    #Ok := "FRK_ConfigDecode"(Text := STRING_TO_WSTRING("FRK_PersistImages".D010.Rows[6].Record.ValueText), Storage := 3, Minimum := 0.0, Maximum := 1000.0, MaxLength := 0, Value := "FRK_ConfigScratch".Value);
    IF NOT #Ok THEN RETURN; END_IF;
    IF NOT "FRK_PersistImages".D010.Rows[7].Used OR "FRK_PersistImages".D010.Rows[7].SchemaVersion <> 4 OR "FRK_PersistImages".D010.Rows[7].ModelCode <> 'MODEL_A' OR "FRK_PersistImages".D010.Rows[7].Record.Scope <> 'StationB.Cell.Gate' OR "FRK_PersistImages".D010.Rows[7].Record.WriteKey <> 'timeout' OR "FRK_PersistImages".D010.Rows[7].Record.Revision <> 1 OR "FRK_PersistImages".D010.Rows[7].Record.Kind <> 0 OR "FRK_PersistImages".D010.Rows[7].Record.ValueType <> 3 THEN RETURN; END_IF;
    #Ok := "FRK_ConfigDecode"(Text := STRING_TO_WSTRING("FRK_PersistImages".D010.Rows[7].Record.ValueText), Storage := 7, Minimum := 1.0, Maximum := 60000.0, MaxLength := 0, Value := "FRK_ConfigScratch".Value);
    IF NOT #Ok THEN RETURN; END_IF;
    IF NOT "FRK_PersistImages".D010.Rows[8].Used OR "FRK_PersistImages".D010.Rows[8].SchemaVersion <> 4 OR "FRK_PersistImages".D010.Rows[8].ModelCode <> 'MODEL_A' OR "FRK_PersistImages".D010.Rows[8].Record.Scope <> 'StationB.Cell.Gate' OR "FRK_PersistImages".D010.Rows[8].Record.WriteKey <> 'preset' OR "FRK_PersistImages".D010.Rows[8].Record.Revision <> 2 OR "FRK_PersistImages".D010.Rows[8].Record.Kind <> 0 OR "FRK_PersistImages".D010.Rows[8].Record.ValueType <> 0 THEN RETURN; END_IF;
    #Ok := "FRK_ConfigDecode"(Text := STRING_TO_WSTRING("FRK_PersistImages".D010.Rows[8].Record.ValueText), Storage := 3, Minimum := 0.0, Maximum := 1000.0, MaxLength := 0, Value := "FRK_ConfigScratch".Value);
    IF NOT #Ok THEN RETURN; END_IF;
    IF NOT "FRK_PersistImages".D010.Rows[9].Used OR "FRK_PersistImages".D010.Rows[9].SchemaVersion <> 4 OR "FRK_PersistImages".D010.Rows[9].ModelCode <> 'MODEL_A' OR "FRK_PersistImages".D010.Rows[9].Record.Scope <> 'StationB.Satellite' OR "FRK_PersistImages".D010.Rows[9].Record.WriteKey <> 'timeout' OR "FRK_PersistImages".D010.Rows[9].Record.Revision <> 1 OR "FRK_PersistImages".D010.Rows[9].Record.Kind <> 0 OR "FRK_PersistImages".D010.Rows[9].Record.ValueType <> 3 THEN RETURN; END_IF;
    #Ok := "FRK_ConfigDecode"(Text := STRING_TO_WSTRING("FRK_PersistImages".D010.Rows[9].Record.ValueText), Storage := 7, Minimum := 1.0, Maximum := 60000.0, MaxLength := 0, Value := "FRK_ConfigScratch".Value);
    IF NOT #Ok THEN RETURN; END_IF;
    IF NOT "FRK_PersistImages".D010.Rows[10].Used OR "FRK_PersistImages".D010.Rows[10].SchemaVersion <> 4 OR "FRK_PersistImages".D010.Rows[10].ModelCode <> 'MODEL_A' OR "FRK_PersistImages".D010.Rows[10].Record.Scope <> 'StationB.Satellite' OR "FRK_PersistImages".D010.Rows[10].Record.WriteKey <> 'preset' OR "FRK_PersistImages".D010.Rows[10].Record.Revision <> 2 OR "FRK_PersistImages".D010.Rows[10].Record.Kind <> 0 OR "FRK_PersistImages".D010.Rows[10].Record.ValueType <> 0 THEN RETURN; END_IF;
    #Ok := "FRK_ConfigDecode"(Text := STRING_TO_WSTRING("FRK_PersistImages".D010.Rows[10].Record.ValueText), Storage := 3, Minimum := 0.0, Maximum := 1000.0, MaxLength := 0, Value := "FRK_ConfigScratch".Value);
    IF NOT #Ok THEN RETURN; END_IF;
    IF NOT "FRK_PersistImages".D010.Rows[11].Used OR "FRK_PersistImages".D010.Rows[11].SchemaVersion <> 4 OR "FRK_PersistImages".D010.Rows[11].ModelCode <> 'MODEL_A' OR "FRK_PersistImages".D010.Rows[11].Record.Scope <> 'StationB.Satellite.Cell' OR "FRK_PersistImages".D010.Rows[11].Record.WriteKey <> 'timeout' OR "FRK_PersistImages".D010.Rows[11].Record.Revision <> 1 OR "FRK_PersistImages".D010.Rows[11].Record.Kind <> 0 OR "FRK_PersistImages".D010.Rows[11].Record.ValueType <> 3 THEN RETURN; END_IF;
    #Ok := "FRK_ConfigDecode"(Text := STRING_TO_WSTRING("FRK_PersistImages".D010.Rows[11].Record.ValueText), Storage := 7, Minimum := 1.0, Maximum := 60000.0, MaxLength := 0, Value := "FRK_ConfigScratch".Value);
    IF NOT #Ok THEN RETURN; END_IF;
    IF NOT "FRK_PersistImages".D010.Rows[12].Used OR "FRK_PersistImages".D010.Rows[12].SchemaVersion <> 4 OR "FRK_PersistImages".D010.Rows[12].ModelCode <> 'MODEL_A' OR "FRK_PersistImages".D010.Rows[12].Record.Scope <> 'StationB.Satellite.Cell' OR "FRK_PersistImages".D010.Rows[12].Record.WriteKey <> 'preset' OR "FRK_PersistImages".D010.Rows[12].Record.Revision <> 2 OR "FRK_PersistImages".D010.Rows[12].Record.Kind <> 0 OR "FRK_PersistImages".D010.Rows[12].Record.ValueType <> 0 THEN RETURN; END_IF;
    #Ok := "FRK_ConfigDecode"(Text := STRING_TO_WSTRING("FRK_PersistImages".D010.Rows[12].Record.ValueText), Storage := 3, Minimum := 0.0, Maximum := 1000.0, MaxLength := 0, Value := "FRK_ConfigScratch".Value);
    IF NOT #Ok THEN RETURN; END_IF;
    IF NOT "FRK_PersistImages".D010.Rows[13].Used OR "FRK_PersistImages".D010.Rows[13].SchemaVersion <> 4 OR "FRK_PersistImages".D010.Rows[13].ModelCode <> 'MODEL_A' OR "FRK_PersistImages".D010.Rows[13].Record.Scope <> 'StationB.Satellite.Cell.Clamp' OR "FRK_PersistImages".D010.Rows[13].Record.WriteKey <> 'timeout' OR "FRK_PersistImages".D010.Rows[13].Record.Revision <> 1 OR "FRK_PersistImages".D010.Rows[13].Record.Kind <> 0 OR "FRK_PersistImages".D010.Rows[13].Record.ValueType <> 3 THEN RETURN; END_IF;
    #Ok := "FRK_ConfigDecode"(Text := STRING_TO_WSTRING("FRK_PersistImages".D010.Rows[13].Record.ValueText), Storage := 7, Minimum := 1.0, Maximum := 60000.0, MaxLength := 0, Value := "FRK_ConfigScratch".Value);
    IF NOT #Ok THEN RETURN; END_IF;
    IF NOT "FRK_PersistImages".D010.Rows[14].Used OR "FRK_PersistImages".D010.Rows[14].SchemaVersion <> 4 OR "FRK_PersistImages".D010.Rows[14].ModelCode <> 'MODEL_A' OR "FRK_PersistImages".D010.Rows[14].Record.Scope <> 'StationB.Satellite.Cell.Clamp' OR "FRK_PersistImages".D010.Rows[14].Record.WriteKey <> 'preset' OR "FRK_PersistImages".D010.Rows[14].Record.Revision <> 2 OR "FRK_PersistImages".D010.Rows[14].Record.Kind <> 0 OR "FRK_PersistImages".D010.Rows[14].Record.ValueType <> 0 THEN RETURN; END_IF;
    #Ok := "FRK_ConfigDecode"(Text := STRING_TO_WSTRING("FRK_PersistImages".D010.Rows[14].Record.ValueText), Storage := 3, Minimum := 0.0, Maximum := 1000.0, MaxLength := 0, Value := "FRK_ConfigScratch".Value);
    IF NOT #Ok THEN RETURN; END_IF;
    IF NOT "FRK_PersistImages".D010.Rows[15].Used OR "FRK_PersistImages".D010.Rows[15].SchemaVersion <> 4 OR "FRK_PersistImages".D010.Rows[15].ModelCode <> 'MODEL_A' OR "FRK_PersistImages".D010.Rows[15].Record.Scope <> 'StationB.Satellite.Cell.Gate' OR "FRK_PersistImages".D010.Rows[15].Record.WriteKey <> 'timeout' OR "FRK_PersistImages".D010.Rows[15].Record.Revision <> 1 OR "FRK_PersistImages".D010.Rows[15].Record.Kind <> 0 OR "FRK_PersistImages".D010.Rows[15].Record.ValueType <> 3 THEN RETURN; END_IF;
    #Ok := "FRK_ConfigDecode"(Text := STRING_TO_WSTRING("FRK_PersistImages".D010.Rows[15].Record.ValueText), Storage := 7, Minimum := 1.0, Maximum := 60000.0, MaxLength := 0, Value := "FRK_ConfigScratch".Value);
    IF NOT #Ok THEN RETURN; END_IF;
    IF NOT "FRK_PersistImages".D010.Rows[16].Used OR "FRK_PersistImages".D010.Rows[16].SchemaVersion <> 4 OR "FRK_PersistImages".D010.Rows[16].ModelCode <> 'MODEL_A' OR "FRK_PersistImages".D010.Rows[16].Record.Scope <> 'StationB.Satellite.Cell.Gate' OR "FRK_PersistImages".D010.Rows[16].Record.WriteKey <> 'preset' OR "FRK_PersistImages".D010.Rows[16].Record.Revision <> 2 OR "FRK_PersistImages".D010.Rows[16].Record.Kind <> 0 OR "FRK_PersistImages".D010.Rows[16].Record.ValueType <> 0 THEN RETURN; END_IF;
    #Ok := "FRK_ConfigDecode"(Text := STRING_TO_WSTRING("FRK_PersistImages".D010.Rows[16].Record.ValueText), Storage := 3, Minimum := 0.0, Maximum := 1000.0, MaxLength := 0, Value := "FRK_ConfigScratch".Value);
    IF NOT #Ok THEN RETURN; END_IF;
    IF NOT "FRK_PersistImages".D010.Rows[17].Used OR "FRK_PersistImages".D010.Rows[17].SchemaVersion <> 4 OR "FRK_PersistImages".D010.Rows[17].ModelCode <> 'MODEL_A' OR "FRK_PersistImages".D010.Rows[17].Record.Scope <> 'StationB.Satellite.Inner' OR "FRK_PersistImages".D010.Rows[17].Record.WriteKey <> 'timeout' OR "FRK_PersistImages".D010.Rows[17].Record.Revision <> 1 OR "FRK_PersistImages".D010.Rows[17].Record.Kind <> 0 OR "FRK_PersistImages".D010.Rows[17].Record.ValueType <> 3 THEN RETURN; END_IF;
    #Ok := "FRK_ConfigDecode"(Text := STRING_TO_WSTRING("FRK_PersistImages".D010.Rows[17].Record.ValueText), Storage := 7, Minimum := 1.0, Maximum := 60000.0, MaxLength := 0, Value := "FRK_ConfigScratch".Value);
    IF NOT #Ok THEN RETURN; END_IF;
    IF NOT "FRK_PersistImages".D010.Rows[18].Used OR "FRK_PersistImages".D010.Rows[18].SchemaVersion <> 4 OR "FRK_PersistImages".D010.Rows[18].ModelCode <> 'MODEL_A' OR "FRK_PersistImages".D010.Rows[18].Record.Scope <> 'StationB.Satellite.Inner' OR "FRK_PersistImages".D010.Rows[18].Record.WriteKey <> 'preset' OR "FRK_PersistImages".D010.Rows[18].Record.Revision <> 2 OR "FRK_PersistImages".D010.Rows[18].Record.Kind <> 0 OR "FRK_PersistImages".D010.Rows[18].Record.ValueType <> 0 THEN RETURN; END_IF;
    #Ok := "FRK_ConfigDecode"(Text := STRING_TO_WSTRING("FRK_PersistImages".D010.Rows[18].Record.ValueText), Storage := 3, Minimum := 0.0, Maximum := 1000.0, MaxLength := 0, Value := "FRK_ConfigScratch".Value);
    IF NOT #Ok THEN RETURN; END_IF;
    IF NOT "FRK_PersistImages".D010.Rows[19].Used OR "FRK_PersistImages".D010.Rows[19].SchemaVersion <> 4 OR "FRK_PersistImages".D010.Rows[19].ModelCode <> 'MODEL_A' OR "FRK_PersistImages".D010.Rows[19].Record.Scope <> 'StationB.Satellite.Inner.Cell' OR "FRK_PersistImages".D010.Rows[19].Record.WriteKey <> 'timeout' OR "FRK_PersistImages".D010.Rows[19].Record.Revision <> 1 OR "FRK_PersistImages".D010.Rows[19].Record.Kind <> 0 OR "FRK_PersistImages".D010.Rows[19].Record.ValueType <> 3 THEN RETURN; END_IF;
    #Ok := "FRK_ConfigDecode"(Text := STRING_TO_WSTRING("FRK_PersistImages".D010.Rows[19].Record.ValueText), Storage := 7, Minimum := 1.0, Maximum := 60000.0, MaxLength := 0, Value := "FRK_ConfigScratch".Value);
    IF NOT #Ok THEN RETURN; END_IF;
    IF NOT "FRK_PersistImages".D010.Rows[20].Used OR "FRK_PersistImages".D010.Rows[20].SchemaVersion <> 4 OR "FRK_PersistImages".D010.Rows[20].ModelCode <> 'MODEL_A' OR "FRK_PersistImages".D010.Rows[20].Record.Scope <> 'StationB.Satellite.Inner.Cell' OR "FRK_PersistImages".D010.Rows[20].Record.WriteKey <> 'preset' OR "FRK_PersistImages".D010.Rows[20].Record.Revision <> 2 OR "FRK_PersistImages".D010.Rows[20].Record.Kind <> 0 OR "FRK_PersistImages".D010.Rows[20].Record.ValueType <> 0 THEN RETURN; END_IF;
    #Ok := "FRK_ConfigDecode"(Text := STRING_TO_WSTRING("FRK_PersistImages".D010.Rows[20].Record.ValueText), Storage := 3, Minimum := 0.0, Maximum := 1000.0, MaxLength := 0, Value := "FRK_ConfigScratch".Value);
    IF NOT #Ok THEN RETURN; END_IF;
    IF NOT "FRK_PersistImages".D010.Rows[21].Used OR "FRK_PersistImages".D010.Rows[21].SchemaVersion <> 4 OR "FRK_PersistImages".D010.Rows[21].ModelCode <> 'MODEL_A' OR "FRK_PersistImages".D010.Rows[21].Record.Scope <> 'StationB.Satellite.Inner.Cell.Clamp' OR "FRK_PersistImages".D010.Rows[21].Record.WriteKey <> 'timeout' OR "FRK_PersistImages".D010.Rows[21].Record.Revision <> 1 OR "FRK_PersistImages".D010.Rows[21].Record.Kind <> 0 OR "FRK_PersistImages".D010.Rows[21].Record.ValueType <> 3 THEN RETURN; END_IF;
    #Ok := "FRK_ConfigDecode"(Text := STRING_TO_WSTRING("FRK_PersistImages".D010.Rows[21].Record.ValueText), Storage := 7, Minimum := 1.0, Maximum := 60000.0, MaxLength := 0, Value := "FRK_ConfigScratch".Value);
    IF NOT #Ok THEN RETURN; END_IF;
    IF NOT "FRK_PersistImages".D010.Rows[22].Used OR "FRK_PersistImages".D010.Rows[22].SchemaVersion <> 4 OR "FRK_PersistImages".D010.Rows[22].ModelCode <> 'MODEL_A' OR "FRK_PersistImages".D010.Rows[22].Record.Scope <> 'StationB.Satellite.Inner.Cell.Clamp' OR "FRK_PersistImages".D010.Rows[22].Record.WriteKey <> 'preset' OR "FRK_PersistImages".D010.Rows[22].Record.Revision <> 2 OR "FRK_PersistImages".D010.Rows[22].Record.Kind <> 0 OR "FRK_PersistImages".D010.Rows[22].Record.ValueType <> 0 THEN RETURN; END_IF;
    #Ok := "FRK_ConfigDecode"(Text := STRING_TO_WSTRING("FRK_PersistImages".D010.Rows[22].Record.ValueText), Storage := 3, Minimum := 0.0, Maximum := 1000.0, MaxLength := 0, Value := "FRK_ConfigScratch".Value);
    IF NOT #Ok THEN RETURN; END_IF;
    IF NOT "FRK_PersistImages".D010.Rows[23].Used OR "FRK_PersistImages".D010.Rows[23].SchemaVersion <> 4 OR "FRK_PersistImages".D010.Rows[23].ModelCode <> 'MODEL_A' OR "FRK_PersistImages".D010.Rows[23].Record.Scope <> 'StationB.Satellite.Inner.Cell.Gate' OR "FRK_PersistImages".D010.Rows[23].Record.WriteKey <> 'timeout' OR "FRK_PersistImages".D010.Rows[23].Record.Revision <> 1 OR "FRK_PersistImages".D010.Rows[23].Record.Kind <> 0 OR "FRK_PersistImages".D010.Rows[23].Record.ValueType <> 3 THEN RETURN; END_IF;
    #Ok := "FRK_ConfigDecode"(Text := STRING_TO_WSTRING("FRK_PersistImages".D010.Rows[23].Record.ValueText), Storage := 7, Minimum := 1.0, Maximum := 60000.0, MaxLength := 0, Value := "FRK_ConfigScratch".Value);
    IF NOT #Ok THEN RETURN; END_IF;
    IF NOT "FRK_PersistImages".D010.Rows[24].Used OR "FRK_PersistImages".D010.Rows[24].SchemaVersion <> 4 OR "FRK_PersistImages".D010.Rows[24].ModelCode <> 'MODEL_A' OR "FRK_PersistImages".D010.Rows[24].Record.Scope <> 'StationB.Satellite.Inner.Cell.Gate' OR "FRK_PersistImages".D010.Rows[24].Record.WriteKey <> 'preset' OR "FRK_PersistImages".D010.Rows[24].Record.Revision <> 2 OR "FRK_PersistImages".D010.Rows[24].Record.Kind <> 0 OR "FRK_PersistImages".D010.Rows[24].Record.ValueType <> 0 THEN RETURN; END_IF;
    #Ok := "FRK_ConfigDecode"(Text := STRING_TO_WSTRING("FRK_PersistImages".D010.Rows[24].Record.ValueText), Storage := 3, Minimum := 0.0, Maximum := 1000.0, MaxLength := 0, Value := "FRK_ConfigScratch".Value);
    IF NOT #Ok THEN RETURN; END_IF;
    #Stored := "FRK_ConfigFind"(Scope := 'StationB', Key := 'timeout', ModelCode := 'MODEL_A');
    IF #Stored = 0 THEN
        FOR #Index := 1 TO 114 DO
            #Reserved := NOT "FRK_ConfigStore".Rows[#Index].Used;
            FOR #Prior := 1 TO 0 DO IF #Targets[#Prior] = #Index THEN #Reserved := FALSE; END_IF; END_FOR;
            IF #Reserved THEN #Stored := #Index; EXIT; END_IF;
        END_FOR;
    END_IF;
    IF #Stored < 1 OR #Stored > 114 THEN RETURN; END_IF;
    #Targets[1] := #Stored;
    #Stored := "FRK_ConfigFind"(Scope := 'StationB', Key := 'preset', ModelCode := 'MODEL_A');
    IF #Stored = 0 THEN
        FOR #Index := 1 TO 114 DO
            #Reserved := NOT "FRK_ConfigStore".Rows[#Index].Used;
            FOR #Prior := 1 TO 1 DO IF #Targets[#Prior] = #Index THEN #Reserved := FALSE; END_IF; END_FOR;
            IF #Reserved THEN #Stored := #Index; EXIT; END_IF;
        END_FOR;
    END_IF;
    IF #Stored < 1 OR #Stored > 114 THEN RETURN; END_IF;
    #Targets[2] := #Stored;
    #Stored := "FRK_ConfigFind"(Scope := 'StationB.Cell', Key := 'timeout', ModelCode := 'MODEL_A');
    IF #Stored = 0 THEN
        FOR #Index := 1 TO 114 DO
            #Reserved := NOT "FRK_ConfigStore".Rows[#Index].Used;
            FOR #Prior := 1 TO 2 DO IF #Targets[#Prior] = #Index THEN #Reserved := FALSE; END_IF; END_FOR;
            IF #Reserved THEN #Stored := #Index; EXIT; END_IF;
        END_FOR;
    END_IF;
    IF #Stored < 1 OR #Stored > 114 THEN RETURN; END_IF;
    #Targets[3] := #Stored;
    #Stored := "FRK_ConfigFind"(Scope := 'StationB.Cell', Key := 'preset', ModelCode := 'MODEL_A');
    IF #Stored = 0 THEN
        FOR #Index := 1 TO 114 DO
            #Reserved := NOT "FRK_ConfigStore".Rows[#Index].Used;
            FOR #Prior := 1 TO 3 DO IF #Targets[#Prior] = #Index THEN #Reserved := FALSE; END_IF; END_FOR;
            IF #Reserved THEN #Stored := #Index; EXIT; END_IF;
        END_FOR;
    END_IF;
    IF #Stored < 1 OR #Stored > 114 THEN RETURN; END_IF;
    #Targets[4] := #Stored;
    #Stored := "FRK_ConfigFind"(Scope := 'StationB.Cell.Clamp', Key := 'timeout', ModelCode := 'MODEL_A');
    IF #Stored = 0 THEN
        FOR #Index := 1 TO 114 DO
            #Reserved := NOT "FRK_ConfigStore".Rows[#Index].Used;
            FOR #Prior := 1 TO 4 DO IF #Targets[#Prior] = #Index THEN #Reserved := FALSE; END_IF; END_FOR;
            IF #Reserved THEN #Stored := #Index; EXIT; END_IF;
        END_FOR;
    END_IF;
    IF #Stored < 1 OR #Stored > 114 THEN RETURN; END_IF;
    #Targets[5] := #Stored;
    #Stored := "FRK_ConfigFind"(Scope := 'StationB.Cell.Clamp', Key := 'preset', ModelCode := 'MODEL_A');
    IF #Stored = 0 THEN
        FOR #Index := 1 TO 114 DO
            #Reserved := NOT "FRK_ConfigStore".Rows[#Index].Used;
            FOR #Prior := 1 TO 5 DO IF #Targets[#Prior] = #Index THEN #Reserved := FALSE; END_IF; END_FOR;
            IF #Reserved THEN #Stored := #Index; EXIT; END_IF;
        END_FOR;
    END_IF;
    IF #Stored < 1 OR #Stored > 114 THEN RETURN; END_IF;
    #Targets[6] := #Stored;
    #Stored := "FRK_ConfigFind"(Scope := 'StationB.Cell.Gate', Key := 'timeout', ModelCode := 'MODEL_A');
    IF #Stored = 0 THEN
        FOR #Index := 1 TO 114 DO
            #Reserved := NOT "FRK_ConfigStore".Rows[#Index].Used;
            FOR #Prior := 1 TO 6 DO IF #Targets[#Prior] = #Index THEN #Reserved := FALSE; END_IF; END_FOR;
            IF #Reserved THEN #Stored := #Index; EXIT; END_IF;
        END_FOR;
    END_IF;
    IF #Stored < 1 OR #Stored > 114 THEN RETURN; END_IF;
    #Targets[7] := #Stored;
    #Stored := "FRK_ConfigFind"(Scope := 'StationB.Cell.Gate', Key := 'preset', ModelCode := 'MODEL_A');
    IF #Stored = 0 THEN
        FOR #Index := 1 TO 114 DO
            #Reserved := NOT "FRK_ConfigStore".Rows[#Index].Used;
            FOR #Prior := 1 TO 7 DO IF #Targets[#Prior] = #Index THEN #Reserved := FALSE; END_IF; END_FOR;
            IF #Reserved THEN #Stored := #Index; EXIT; END_IF;
        END_FOR;
    END_IF;
    IF #Stored < 1 OR #Stored > 114 THEN RETURN; END_IF;
    #Targets[8] := #Stored;
    #Stored := "FRK_ConfigFind"(Scope := 'StationB.Satellite', Key := 'timeout', ModelCode := 'MODEL_A');
    IF #Stored = 0 THEN
        FOR #Index := 1 TO 114 DO
            #Reserved := NOT "FRK_ConfigStore".Rows[#Index].Used;
            FOR #Prior := 1 TO 8 DO IF #Targets[#Prior] = #Index THEN #Reserved := FALSE; END_IF; END_FOR;
            IF #Reserved THEN #Stored := #Index; EXIT; END_IF;
        END_FOR;
    END_IF;
    IF #Stored < 1 OR #Stored > 114 THEN RETURN; END_IF;
    #Targets[9] := #Stored;
    #Stored := "FRK_ConfigFind"(Scope := 'StationB.Satellite', Key := 'preset', ModelCode := 'MODEL_A');
    IF #Stored = 0 THEN
        FOR #Index := 1 TO 114 DO
            #Reserved := NOT "FRK_ConfigStore".Rows[#Index].Used;
            FOR #Prior := 1 TO 9 DO IF #Targets[#Prior] = #Index THEN #Reserved := FALSE; END_IF; END_FOR;
            IF #Reserved THEN #Stored := #Index; EXIT; END_IF;
        END_FOR;
    END_IF;
    IF #Stored < 1 OR #Stored > 114 THEN RETURN; END_IF;
    #Targets[10] := #Stored;
    #Stored := "FRK_ConfigFind"(Scope := 'StationB.Satellite.Cell', Key := 'timeout', ModelCode := 'MODEL_A');
    IF #Stored = 0 THEN
        FOR #Index := 1 TO 114 DO
            #Reserved := NOT "FRK_ConfigStore".Rows[#Index].Used;
            FOR #Prior := 1 TO 10 DO IF #Targets[#Prior] = #Index THEN #Reserved := FALSE; END_IF; END_FOR;
            IF #Reserved THEN #Stored := #Index; EXIT; END_IF;
        END_FOR;
    END_IF;
    IF #Stored < 1 OR #Stored > 114 THEN RETURN; END_IF;
    #Targets[11] := #Stored;
    #Stored := "FRK_ConfigFind"(Scope := 'StationB.Satellite.Cell', Key := 'preset', ModelCode := 'MODEL_A');
    IF #Stored = 0 THEN
        FOR #Index := 1 TO 114 DO
            #Reserved := NOT "FRK_ConfigStore".Rows[#Index].Used;
            FOR #Prior := 1 TO 11 DO IF #Targets[#Prior] = #Index THEN #Reserved := FALSE; END_IF; END_FOR;
            IF #Reserved THEN #Stored := #Index; EXIT; END_IF;
        END_FOR;
    END_IF;
    IF #Stored < 1 OR #Stored > 114 THEN RETURN; END_IF;
    #Targets[12] := #Stored;
    #Stored := "FRK_ConfigFind"(Scope := 'StationB.Satellite.Cell.Clamp', Key := 'timeout', ModelCode := 'MODEL_A');
    IF #Stored = 0 THEN
        FOR #Index := 1 TO 114 DO
            #Reserved := NOT "FRK_ConfigStore".Rows[#Index].Used;
            FOR #Prior := 1 TO 12 DO IF #Targets[#Prior] = #Index THEN #Reserved := FALSE; END_IF; END_FOR;
            IF #Reserved THEN #Stored := #Index; EXIT; END_IF;
        END_FOR;
    END_IF;
    IF #Stored < 1 OR #Stored > 114 THEN RETURN; END_IF;
    #Targets[13] := #Stored;
    #Stored := "FRK_ConfigFind"(Scope := 'StationB.Satellite.Cell.Clamp', Key := 'preset', ModelCode := 'MODEL_A');
    IF #Stored = 0 THEN
        FOR #Index := 1 TO 114 DO
            #Reserved := NOT "FRK_ConfigStore".Rows[#Index].Used;
            FOR #Prior := 1 TO 13 DO IF #Targets[#Prior] = #Index THEN #Reserved := FALSE; END_IF; END_FOR;
            IF #Reserved THEN #Stored := #Index; EXIT; END_IF;
        END_FOR;
    END_IF;
    IF #Stored < 1 OR #Stored > 114 THEN RETURN; END_IF;
    #Targets[14] := #Stored;
    #Stored := "FRK_ConfigFind"(Scope := 'StationB.Satellite.Cell.Gate', Key := 'timeout', ModelCode := 'MODEL_A');
    IF #Stored = 0 THEN
        FOR #Index := 1 TO 114 DO
            #Reserved := NOT "FRK_ConfigStore".Rows[#Index].Used;
            FOR #Prior := 1 TO 14 DO IF #Targets[#Prior] = #Index THEN #Reserved := FALSE; END_IF; END_FOR;
            IF #Reserved THEN #Stored := #Index; EXIT; END_IF;
        END_FOR;
    END_IF;
    IF #Stored < 1 OR #Stored > 114 THEN RETURN; END_IF;
    #Targets[15] := #Stored;
    #Stored := "FRK_ConfigFind"(Scope := 'StationB.Satellite.Cell.Gate', Key := 'preset', ModelCode := 'MODEL_A');
    IF #Stored = 0 THEN
        FOR #Index := 1 TO 114 DO
            #Reserved := NOT "FRK_ConfigStore".Rows[#Index].Used;
            FOR #Prior := 1 TO 15 DO IF #Targets[#Prior] = #Index THEN #Reserved := FALSE; END_IF; END_FOR;
            IF #Reserved THEN #Stored := #Index; EXIT; END_IF;
        END_FOR;
    END_IF;
    IF #Stored < 1 OR #Stored > 114 THEN RETURN; END_IF;
    #Targets[16] := #Stored;
    #Stored := "FRK_ConfigFind"(Scope := 'StationB.Satellite.Inner', Key := 'timeout', ModelCode := 'MODEL_A');
    IF #Stored = 0 THEN
        FOR #Index := 1 TO 114 DO
            #Reserved := NOT "FRK_ConfigStore".Rows[#Index].Used;
            FOR #Prior := 1 TO 16 DO IF #Targets[#Prior] = #Index THEN #Reserved := FALSE; END_IF; END_FOR;
            IF #Reserved THEN #Stored := #Index; EXIT; END_IF;
        END_FOR;
    END_IF;
    IF #Stored < 1 OR #Stored > 114 THEN RETURN; END_IF;
    #Targets[17] := #Stored;
    #Stored := "FRK_ConfigFind"(Scope := 'StationB.Satellite.Inner', Key := 'preset', ModelCode := 'MODEL_A');
    IF #Stored = 0 THEN
        FOR #Index := 1 TO 114 DO
            #Reserved := NOT "FRK_ConfigStore".Rows[#Index].Used;
            FOR #Prior := 1 TO 17 DO IF #Targets[#Prior] = #Index THEN #Reserved := FALSE; END_IF; END_FOR;
            IF #Reserved THEN #Stored := #Index; EXIT; END_IF;
        END_FOR;
    END_IF;
    IF #Stored < 1 OR #Stored > 114 THEN RETURN; END_IF;
    #Targets[18] := #Stored;
    #Stored := "FRK_ConfigFind"(Scope := 'StationB.Satellite.Inner.Cell', Key := 'timeout', ModelCode := 'MODEL_A');
    IF #Stored = 0 THEN
        FOR #Index := 1 TO 114 DO
            #Reserved := NOT "FRK_ConfigStore".Rows[#Index].Used;
            FOR #Prior := 1 TO 18 DO IF #Targets[#Prior] = #Index THEN #Reserved := FALSE; END_IF; END_FOR;
            IF #Reserved THEN #Stored := #Index; EXIT; END_IF;
        END_FOR;
    END_IF;
    IF #Stored < 1 OR #Stored > 114 THEN RETURN; END_IF;
    #Targets[19] := #Stored;
    #Stored := "FRK_ConfigFind"(Scope := 'StationB.Satellite.Inner.Cell', Key := 'preset', ModelCode := 'MODEL_A');
    IF #Stored = 0 THEN
        FOR #Index := 1 TO 114 DO
            #Reserved := NOT "FRK_ConfigStore".Rows[#Index].Used;
            FOR #Prior := 1 TO 19 DO IF #Targets[#Prior] = #Index THEN #Reserved := FALSE; END_IF; END_FOR;
            IF #Reserved THEN #Stored := #Index; EXIT; END_IF;
        END_FOR;
    END_IF;
    IF #Stored < 1 OR #Stored > 114 THEN RETURN; END_IF;
    #Targets[20] := #Stored;
    #Stored := "FRK_ConfigFind"(Scope := 'StationB.Satellite.Inner.Cell.Clamp', Key := 'timeout', ModelCode := 'MODEL_A');
    IF #Stored = 0 THEN
        FOR #Index := 1 TO 114 DO
            #Reserved := NOT "FRK_ConfigStore".Rows[#Index].Used;
            FOR #Prior := 1 TO 20 DO IF #Targets[#Prior] = #Index THEN #Reserved := FALSE; END_IF; END_FOR;
            IF #Reserved THEN #Stored := #Index; EXIT; END_IF;
        END_FOR;
    END_IF;
    IF #Stored < 1 OR #Stored > 114 THEN RETURN; END_IF;
    #Targets[21] := #Stored;
    #Stored := "FRK_ConfigFind"(Scope := 'StationB.Satellite.Inner.Cell.Clamp', Key := 'preset', ModelCode := 'MODEL_A');
    IF #Stored = 0 THEN
        FOR #Index := 1 TO 114 DO
            #Reserved := NOT "FRK_ConfigStore".Rows[#Index].Used;
            FOR #Prior := 1 TO 21 DO IF #Targets[#Prior] = #Index THEN #Reserved := FALSE; END_IF; END_FOR;
            IF #Reserved THEN #Stored := #Index; EXIT; END_IF;
        END_FOR;
    END_IF;
    IF #Stored < 1 OR #Stored > 114 THEN RETURN; END_IF;
    #Targets[22] := #Stored;
    #Stored := "FRK_ConfigFind"(Scope := 'StationB.Satellite.Inner.Cell.Gate', Key := 'timeout', ModelCode := 'MODEL_A');
    IF #Stored = 0 THEN
        FOR #Index := 1 TO 114 DO
            #Reserved := NOT "FRK_ConfigStore".Rows[#Index].Used;
            FOR #Prior := 1 TO 22 DO IF #Targets[#Prior] = #Index THEN #Reserved := FALSE; END_IF; END_FOR;
            IF #Reserved THEN #Stored := #Index; EXIT; END_IF;
        END_FOR;
    END_IF;
    IF #Stored < 1 OR #Stored > 114 THEN RETURN; END_IF;
    #Targets[23] := #Stored;
    #Stored := "FRK_ConfigFind"(Scope := 'StationB.Satellite.Inner.Cell.Gate', Key := 'preset', ModelCode := 'MODEL_A');
    IF #Stored = 0 THEN
        FOR #Index := 1 TO 114 DO
            #Reserved := NOT "FRK_ConfigStore".Rows[#Index].Used;
            FOR #Prior := 1 TO 23 DO IF #Targets[#Prior] = #Index THEN #Reserved := FALSE; END_IF; END_FOR;
            IF #Reserved THEN #Stored := #Index; EXIT; END_IF;
        END_FOR;
    END_IF;
    IF #Stored < 1 OR #Stored > 114 THEN RETURN; END_IF;
    #Targets[24] := #Stored;
    "FRK_ConfigStore".Rows[#Targets[1]] := "FRK_PersistImages".D010.Rows[1];
    "FRK_ConfigStore".Rows[#Targets[2]] := "FRK_PersistImages".D010.Rows[2];
    "FRK_ConfigStore".Rows[#Targets[3]] := "FRK_PersistImages".D010.Rows[3];
    "FRK_ConfigStore".Rows[#Targets[4]] := "FRK_PersistImages".D010.Rows[4];
    "FRK_ConfigStore".Rows[#Targets[5]] := "FRK_PersistImages".D010.Rows[5];
    "FRK_ConfigStore".Rows[#Targets[6]] := "FRK_PersistImages".D010.Rows[6];
    "FRK_ConfigStore".Rows[#Targets[7]] := "FRK_PersistImages".D010.Rows[7];
    "FRK_ConfigStore".Rows[#Targets[8]] := "FRK_PersistImages".D010.Rows[8];
    "FRK_ConfigStore".Rows[#Targets[9]] := "FRK_PersistImages".D010.Rows[9];
    "FRK_ConfigStore".Rows[#Targets[10]] := "FRK_PersistImages".D010.Rows[10];
    "FRK_ConfigStore".Rows[#Targets[11]] := "FRK_PersistImages".D010.Rows[11];
    "FRK_ConfigStore".Rows[#Targets[12]] := "FRK_PersistImages".D010.Rows[12];
    "FRK_ConfigStore".Rows[#Targets[13]] := "FRK_PersistImages".D010.Rows[13];
    "FRK_ConfigStore".Rows[#Targets[14]] := "FRK_PersistImages".D010.Rows[14];
    "FRK_ConfigStore".Rows[#Targets[15]] := "FRK_PersistImages".D010.Rows[15];
    "FRK_ConfigStore".Rows[#Targets[16]] := "FRK_PersistImages".D010.Rows[16];
    "FRK_ConfigStore".Rows[#Targets[17]] := "FRK_PersistImages".D010.Rows[17];
    "FRK_ConfigStore".Rows[#Targets[18]] := "FRK_PersistImages".D010.Rows[18];
    "FRK_ConfigStore".Rows[#Targets[19]] := "FRK_PersistImages".D010.Rows[19];
    "FRK_ConfigStore".Rows[#Targets[20]] := "FRK_PersistImages".D010.Rows[20];
    "FRK_ConfigStore".Rows[#Targets[21]] := "FRK_PersistImages".D010.Rows[21];
    "FRK_ConfigStore".Rows[#Targets[22]] := "FRK_PersistImages".D010.Rows[22];
    "FRK_ConfigStore".Rows[#Targets[23]] := "FRK_PersistImages".D010.Rows[23];
    "FRK_ConfigStore".Rows[#Targets[24]] := "FRK_PersistImages".D010.Rows[24];
    "FRK_ConfigStore".SchemaVersion := 1;
    #FRK_DocApply_D010 := TRUE;
END_FUNCTION
FUNCTION "FRK_DocCapture_D011" : Bool
{ S7_Optimized_Access := 'TRUE' }
VERSION : 0.1
VAR_IN_OUT
    Length : DInt;
END_VAR
VAR_TEMP
    Index : Int;
    Stored : Int;
    Position : DInt;
    NativeResult : Int;
    Ok : Bool;
    Targets : Array[1..24] of Int;
    Prior : Int;
    Reserved : Bool;
END_VAR
BEGIN
    #FRK_DocCapture_D011 := FALSE;
    "FRK_PersistImages".D011.SchemaVersion := 1; "FRK_PersistImages".D011.Scope := 'StationB';
    "FRK_PersistImages".D011.Kind := 0;
    "FRK_PersistImages".D011.ModelCode := 'MODEL_B';
    "FRK_PersistImages".D011.ActiveModel := "FRK_ConfigStore".ActiveModels[2];
    "FRK_PersistImages".D011.Count := 24;
    #Stored := "FRK_ConfigFind"(Scope := 'StationB', Key := 'timeout', ModelCode := 'MODEL_B');
    IF #Stored = 0 THEN RETURN; END_IF;
    "FRK_PersistImages".D011.Rows[1] := "FRK_ConfigStore".Rows[#Stored];
    #Stored := "FRK_ConfigFind"(Scope := 'StationB', Key := 'preset', ModelCode := 'MODEL_B');
    IF #Stored = 0 THEN RETURN; END_IF;
    "FRK_PersistImages".D011.Rows[2] := "FRK_ConfigStore".Rows[#Stored];
    #Stored := "FRK_ConfigFind"(Scope := 'StationB.Cell', Key := 'timeout', ModelCode := 'MODEL_B');
    IF #Stored = 0 THEN RETURN; END_IF;
    "FRK_PersistImages".D011.Rows[3] := "FRK_ConfigStore".Rows[#Stored];
    #Stored := "FRK_ConfigFind"(Scope := 'StationB.Cell', Key := 'preset', ModelCode := 'MODEL_B');
    IF #Stored = 0 THEN RETURN; END_IF;
    "FRK_PersistImages".D011.Rows[4] := "FRK_ConfigStore".Rows[#Stored];
    #Stored := "FRK_ConfigFind"(Scope := 'StationB.Cell.Clamp', Key := 'timeout', ModelCode := 'MODEL_B');
    IF #Stored = 0 THEN RETURN; END_IF;
    "FRK_PersistImages".D011.Rows[5] := "FRK_ConfigStore".Rows[#Stored];
    #Stored := "FRK_ConfigFind"(Scope := 'StationB.Cell.Clamp', Key := 'preset', ModelCode := 'MODEL_B');
    IF #Stored = 0 THEN RETURN; END_IF;
    "FRK_PersistImages".D011.Rows[6] := "FRK_ConfigStore".Rows[#Stored];
    #Stored := "FRK_ConfigFind"(Scope := 'StationB.Cell.Gate', Key := 'timeout', ModelCode := 'MODEL_B');
    IF #Stored = 0 THEN RETURN; END_IF;
    "FRK_PersistImages".D011.Rows[7] := "FRK_ConfigStore".Rows[#Stored];
    #Stored := "FRK_ConfigFind"(Scope := 'StationB.Cell.Gate', Key := 'preset', ModelCode := 'MODEL_B');
    IF #Stored = 0 THEN RETURN; END_IF;
    "FRK_PersistImages".D011.Rows[8] := "FRK_ConfigStore".Rows[#Stored];
    #Stored := "FRK_ConfigFind"(Scope := 'StationB.Satellite', Key := 'timeout', ModelCode := 'MODEL_B');
    IF #Stored = 0 THEN RETURN; END_IF;
    "FRK_PersistImages".D011.Rows[9] := "FRK_ConfigStore".Rows[#Stored];
    #Stored := "FRK_ConfigFind"(Scope := 'StationB.Satellite', Key := 'preset', ModelCode := 'MODEL_B');
    IF #Stored = 0 THEN RETURN; END_IF;
    "FRK_PersistImages".D011.Rows[10] := "FRK_ConfigStore".Rows[#Stored];
    #Stored := "FRK_ConfigFind"(Scope := 'StationB.Satellite.Cell', Key := 'timeout', ModelCode := 'MODEL_B');
    IF #Stored = 0 THEN RETURN; END_IF;
    "FRK_PersistImages".D011.Rows[11] := "FRK_ConfigStore".Rows[#Stored];
    #Stored := "FRK_ConfigFind"(Scope := 'StationB.Satellite.Cell', Key := 'preset', ModelCode := 'MODEL_B');
    IF #Stored = 0 THEN RETURN; END_IF;
    "FRK_PersistImages".D011.Rows[12] := "FRK_ConfigStore".Rows[#Stored];
    #Stored := "FRK_ConfigFind"(Scope := 'StationB.Satellite.Cell.Clamp', Key := 'timeout', ModelCode := 'MODEL_B');
    IF #Stored = 0 THEN RETURN; END_IF;
    "FRK_PersistImages".D011.Rows[13] := "FRK_ConfigStore".Rows[#Stored];
    #Stored := "FRK_ConfigFind"(Scope := 'StationB.Satellite.Cell.Clamp', Key := 'preset', ModelCode := 'MODEL_B');
    IF #Stored = 0 THEN RETURN; END_IF;
    "FRK_PersistImages".D011.Rows[14] := "FRK_ConfigStore".Rows[#Stored];
    #Stored := "FRK_ConfigFind"(Scope := 'StationB.Satellite.Cell.Gate', Key := 'timeout', ModelCode := 'MODEL_B');
    IF #Stored = 0 THEN RETURN; END_IF;
    "FRK_PersistImages".D011.Rows[15] := "FRK_ConfigStore".Rows[#Stored];
    #Stored := "FRK_ConfigFind"(Scope := 'StationB.Satellite.Cell.Gate', Key := 'preset', ModelCode := 'MODEL_B');
    IF #Stored = 0 THEN RETURN; END_IF;
    "FRK_PersistImages".D011.Rows[16] := "FRK_ConfigStore".Rows[#Stored];
    #Stored := "FRK_ConfigFind"(Scope := 'StationB.Satellite.Inner', Key := 'timeout', ModelCode := 'MODEL_B');
    IF #Stored = 0 THEN RETURN; END_IF;
    "FRK_PersistImages".D011.Rows[17] := "FRK_ConfigStore".Rows[#Stored];
    #Stored := "FRK_ConfigFind"(Scope := 'StationB.Satellite.Inner', Key := 'preset', ModelCode := 'MODEL_B');
    IF #Stored = 0 THEN RETURN; END_IF;
    "FRK_PersistImages".D011.Rows[18] := "FRK_ConfigStore".Rows[#Stored];
    #Stored := "FRK_ConfigFind"(Scope := 'StationB.Satellite.Inner.Cell', Key := 'timeout', ModelCode := 'MODEL_B');
    IF #Stored = 0 THEN RETURN; END_IF;
    "FRK_PersistImages".D011.Rows[19] := "FRK_ConfigStore".Rows[#Stored];
    #Stored := "FRK_ConfigFind"(Scope := 'StationB.Satellite.Inner.Cell', Key := 'preset', ModelCode := 'MODEL_B');
    IF #Stored = 0 THEN RETURN; END_IF;
    "FRK_PersistImages".D011.Rows[20] := "FRK_ConfigStore".Rows[#Stored];
    #Stored := "FRK_ConfigFind"(Scope := 'StationB.Satellite.Inner.Cell.Clamp', Key := 'timeout', ModelCode := 'MODEL_B');
    IF #Stored = 0 THEN RETURN; END_IF;
    "FRK_PersistImages".D011.Rows[21] := "FRK_ConfigStore".Rows[#Stored];
    #Stored := "FRK_ConfigFind"(Scope := 'StationB.Satellite.Inner.Cell.Clamp', Key := 'preset', ModelCode := 'MODEL_B');
    IF #Stored = 0 THEN RETURN; END_IF;
    "FRK_PersistImages".D011.Rows[22] := "FRK_ConfigStore".Rows[#Stored];
    #Stored := "FRK_ConfigFind"(Scope := 'StationB.Satellite.Inner.Cell.Gate', Key := 'timeout', ModelCode := 'MODEL_B');
    IF #Stored = 0 THEN RETURN; END_IF;
    "FRK_PersistImages".D011.Rows[23] := "FRK_ConfigStore".Rows[#Stored];
    #Stored := "FRK_ConfigFind"(Scope := 'StationB.Satellite.Inner.Cell.Gate', Key := 'preset', ModelCode := 'MODEL_B');
    IF #Stored = 0 THEN RETURN; END_IF;
    "FRK_PersistImages".D011.Rows[24] := "FRK_ConfigStore".Rows[#Stored];
    FOR #Index := 0 TO 11401 DO "FRK_PersistBuffers".D011Data[#Index] := BYTE#0; END_FOR;
    #Position := 24;
    #NativeResult := Serialize(SRC_VARIABLE := "FRK_PersistImages".D011, DEST_ARRAY => "FRK_PersistBuffers".D011Data, POS := #Position);
    IF #NativeResult <> 0 OR #Position < 24 OR #Position > 11402 THEN RETURN; END_IF;
    #Length := #Position - 24;
    #FRK_DocCapture_D011 := TRUE;
END_FUNCTION
FUNCTION "FRK_DocApply_D011" : Bool
{ S7_Optimized_Access := 'TRUE' }
VERSION : 0.1
VAR_TEMP
    Index : Int;
    Stored : Int;
    Position : DInt;
    NativeResult : Int;
    Ok : Bool;
    Targets : Array[1..24] of Int;
    Prior : Int;
    Reserved : Bool;
END_VAR
BEGIN
    #FRK_DocApply_D011 := FALSE;
    #Position := 24;
    #NativeResult := Deserialize(SRC_ARRAY := "FRK_PersistBuffers".D011Data, DEST_VARIABLE => "FRK_PersistImages".D011, POS := #Position);
    IF #NativeResult <> 0 OR #Position <> 24 + UDINT_TO_DINT("FRK_PersistConsumers".Rows[11].Result.Length) THEN RETURN; END_IF;
    IF "FRK_PersistImages".D011.SchemaVersion <> 1 OR "FRK_PersistImages".D011.Scope <> 'StationB' THEN RETURN; END_IF;
    IF "FRK_PersistImages".D011.Kind <> 0 OR "FRK_PersistImages".D011.ModelCode <> 'MODEL_B' OR "FRK_PersistImages".D011.Count <> 24 THEN RETURN; END_IF;
    IF "FRK_PersistImages".D011.ActiveModel <> 'MODEL_A' AND "FRK_PersistImages".D011.ActiveModel <> 'MODEL_B' THEN RETURN; END_IF;
    IF NOT "FRK_PersistImages".D011.Rows[1].Used OR "FRK_PersistImages".D011.Rows[1].SchemaVersion <> 4 OR "FRK_PersistImages".D011.Rows[1].ModelCode <> 'MODEL_B' OR "FRK_PersistImages".D011.Rows[1].Record.Scope <> 'StationB' OR "FRK_PersistImages".D011.Rows[1].Record.WriteKey <> 'timeout' OR "FRK_PersistImages".D011.Rows[1].Record.Revision <> 1 OR "FRK_PersistImages".D011.Rows[1].Record.Kind <> 0 OR "FRK_PersistImages".D011.Rows[1].Record.ValueType <> 3 THEN RETURN; END_IF;
    #Ok := "FRK_ConfigDecode"(Text := STRING_TO_WSTRING("FRK_PersistImages".D011.Rows[1].Record.ValueText), Storage := 7, Minimum := 1.0, Maximum := 60000.0, MaxLength := 0, Value := "FRK_ConfigScratch".Value);
    IF NOT #Ok THEN RETURN; END_IF;
    IF NOT "FRK_PersistImages".D011.Rows[2].Used OR "FRK_PersistImages".D011.Rows[2].SchemaVersion <> 4 OR "FRK_PersistImages".D011.Rows[2].ModelCode <> 'MODEL_B' OR "FRK_PersistImages".D011.Rows[2].Record.Scope <> 'StationB' OR "FRK_PersistImages".D011.Rows[2].Record.WriteKey <> 'preset' OR "FRK_PersistImages".D011.Rows[2].Record.Revision <> 2 OR "FRK_PersistImages".D011.Rows[2].Record.Kind <> 0 OR "FRK_PersistImages".D011.Rows[2].Record.ValueType <> 0 THEN RETURN; END_IF;
    #Ok := "FRK_ConfigDecode"(Text := STRING_TO_WSTRING("FRK_PersistImages".D011.Rows[2].Record.ValueText), Storage := 3, Minimum := 0.0, Maximum := 1000.0, MaxLength := 0, Value := "FRK_ConfigScratch".Value);
    IF NOT #Ok THEN RETURN; END_IF;
    IF NOT "FRK_PersistImages".D011.Rows[3].Used OR "FRK_PersistImages".D011.Rows[3].SchemaVersion <> 4 OR "FRK_PersistImages".D011.Rows[3].ModelCode <> 'MODEL_B' OR "FRK_PersistImages".D011.Rows[3].Record.Scope <> 'StationB.Cell' OR "FRK_PersistImages".D011.Rows[3].Record.WriteKey <> 'timeout' OR "FRK_PersistImages".D011.Rows[3].Record.Revision <> 1 OR "FRK_PersistImages".D011.Rows[3].Record.Kind <> 0 OR "FRK_PersistImages".D011.Rows[3].Record.ValueType <> 3 THEN RETURN; END_IF;
    #Ok := "FRK_ConfigDecode"(Text := STRING_TO_WSTRING("FRK_PersistImages".D011.Rows[3].Record.ValueText), Storage := 7, Minimum := 1.0, Maximum := 60000.0, MaxLength := 0, Value := "FRK_ConfigScratch".Value);
    IF NOT #Ok THEN RETURN; END_IF;
    IF NOT "FRK_PersistImages".D011.Rows[4].Used OR "FRK_PersistImages".D011.Rows[4].SchemaVersion <> 4 OR "FRK_PersistImages".D011.Rows[4].ModelCode <> 'MODEL_B' OR "FRK_PersistImages".D011.Rows[4].Record.Scope <> 'StationB.Cell' OR "FRK_PersistImages".D011.Rows[4].Record.WriteKey <> 'preset' OR "FRK_PersistImages".D011.Rows[4].Record.Revision <> 2 OR "FRK_PersistImages".D011.Rows[4].Record.Kind <> 0 OR "FRK_PersistImages".D011.Rows[4].Record.ValueType <> 0 THEN RETURN; END_IF;
    #Ok := "FRK_ConfigDecode"(Text := STRING_TO_WSTRING("FRK_PersistImages".D011.Rows[4].Record.ValueText), Storage := 3, Minimum := 0.0, Maximum := 1000.0, MaxLength := 0, Value := "FRK_ConfigScratch".Value);
    IF NOT #Ok THEN RETURN; END_IF;
    IF NOT "FRK_PersistImages".D011.Rows[5].Used OR "FRK_PersistImages".D011.Rows[5].SchemaVersion <> 4 OR "FRK_PersistImages".D011.Rows[5].ModelCode <> 'MODEL_B' OR "FRK_PersistImages".D011.Rows[5].Record.Scope <> 'StationB.Cell.Clamp' OR "FRK_PersistImages".D011.Rows[5].Record.WriteKey <> 'timeout' OR "FRK_PersistImages".D011.Rows[5].Record.Revision <> 1 OR "FRK_PersistImages".D011.Rows[5].Record.Kind <> 0 OR "FRK_PersistImages".D011.Rows[5].Record.ValueType <> 3 THEN RETURN; END_IF;
    #Ok := "FRK_ConfigDecode"(Text := STRING_TO_WSTRING("FRK_PersistImages".D011.Rows[5].Record.ValueText), Storage := 7, Minimum := 1.0, Maximum := 60000.0, MaxLength := 0, Value := "FRK_ConfigScratch".Value);
    IF NOT #Ok THEN RETURN; END_IF;
    IF NOT "FRK_PersistImages".D011.Rows[6].Used OR "FRK_PersistImages".D011.Rows[6].SchemaVersion <> 4 OR "FRK_PersistImages".D011.Rows[6].ModelCode <> 'MODEL_B' OR "FRK_PersistImages".D011.Rows[6].Record.Scope <> 'StationB.Cell.Clamp' OR "FRK_PersistImages".D011.Rows[6].Record.WriteKey <> 'preset' OR "FRK_PersistImages".D011.Rows[6].Record.Revision <> 2 OR "FRK_PersistImages".D011.Rows[6].Record.Kind <> 0 OR "FRK_PersistImages".D011.Rows[6].Record.ValueType <> 0 THEN RETURN; END_IF;
    #Ok := "FRK_ConfigDecode"(Text := STRING_TO_WSTRING("FRK_PersistImages".D011.Rows[6].Record.ValueText), Storage := 3, Minimum := 0.0, Maximum := 1000.0, MaxLength := 0, Value := "FRK_ConfigScratch".Value);
    IF NOT #Ok THEN RETURN; END_IF;
    IF NOT "FRK_PersistImages".D011.Rows[7].Used OR "FRK_PersistImages".D011.Rows[7].SchemaVersion <> 4 OR "FRK_PersistImages".D011.Rows[7].ModelCode <> 'MODEL_B' OR "FRK_PersistImages".D011.Rows[7].Record.Scope <> 'StationB.Cell.Gate' OR "FRK_PersistImages".D011.Rows[7].Record.WriteKey <> 'timeout' OR "FRK_PersistImages".D011.Rows[7].Record.Revision <> 1 OR "FRK_PersistImages".D011.Rows[7].Record.Kind <> 0 OR "FRK_PersistImages".D011.Rows[7].Record.ValueType <> 3 THEN RETURN; END_IF;
    #Ok := "FRK_ConfigDecode"(Text := STRING_TO_WSTRING("FRK_PersistImages".D011.Rows[7].Record.ValueText), Storage := 7, Minimum := 1.0, Maximum := 60000.0, MaxLength := 0, Value := "FRK_ConfigScratch".Value);
    IF NOT #Ok THEN RETURN; END_IF;
    IF NOT "FRK_PersistImages".D011.Rows[8].Used OR "FRK_PersistImages".D011.Rows[8].SchemaVersion <> 4 OR "FRK_PersistImages".D011.Rows[8].ModelCode <> 'MODEL_B' OR "FRK_PersistImages".D011.Rows[8].Record.Scope <> 'StationB.Cell.Gate' OR "FRK_PersistImages".D011.Rows[8].Record.WriteKey <> 'preset' OR "FRK_PersistImages".D011.Rows[8].Record.Revision <> 2 OR "FRK_PersistImages".D011.Rows[8].Record.Kind <> 0 OR "FRK_PersistImages".D011.Rows[8].Record.ValueType <> 0 THEN RETURN; END_IF;
    #Ok := "FRK_ConfigDecode"(Text := STRING_TO_WSTRING("FRK_PersistImages".D011.Rows[8].Record.ValueText), Storage := 3, Minimum := 0.0, Maximum := 1000.0, MaxLength := 0, Value := "FRK_ConfigScratch".Value);
    IF NOT #Ok THEN RETURN; END_IF;
    IF NOT "FRK_PersistImages".D011.Rows[9].Used OR "FRK_PersistImages".D011.Rows[9].SchemaVersion <> 4 OR "FRK_PersistImages".D011.Rows[9].ModelCode <> 'MODEL_B' OR "FRK_PersistImages".D011.Rows[9].Record.Scope <> 'StationB.Satellite' OR "FRK_PersistImages".D011.Rows[9].Record.WriteKey <> 'timeout' OR "FRK_PersistImages".D011.Rows[9].Record.Revision <> 1 OR "FRK_PersistImages".D011.Rows[9].Record.Kind <> 0 OR "FRK_PersistImages".D011.Rows[9].Record.ValueType <> 3 THEN RETURN; END_IF;
    #Ok := "FRK_ConfigDecode"(Text := STRING_TO_WSTRING("FRK_PersistImages".D011.Rows[9].Record.ValueText), Storage := 7, Minimum := 1.0, Maximum := 60000.0, MaxLength := 0, Value := "FRK_ConfigScratch".Value);
    IF NOT #Ok THEN RETURN; END_IF;
    IF NOT "FRK_PersistImages".D011.Rows[10].Used OR "FRK_PersistImages".D011.Rows[10].SchemaVersion <> 4 OR "FRK_PersistImages".D011.Rows[10].ModelCode <> 'MODEL_B' OR "FRK_PersistImages".D011.Rows[10].Record.Scope <> 'StationB.Satellite' OR "FRK_PersistImages".D011.Rows[10].Record.WriteKey <> 'preset' OR "FRK_PersistImages".D011.Rows[10].Record.Revision <> 2 OR "FRK_PersistImages".D011.Rows[10].Record.Kind <> 0 OR "FRK_PersistImages".D011.Rows[10].Record.ValueType <> 0 THEN RETURN; END_IF;
    #Ok := "FRK_ConfigDecode"(Text := STRING_TO_WSTRING("FRK_PersistImages".D011.Rows[10].Record.ValueText), Storage := 3, Minimum := 0.0, Maximum := 1000.0, MaxLength := 0, Value := "FRK_ConfigScratch".Value);
    IF NOT #Ok THEN RETURN; END_IF;
    IF NOT "FRK_PersistImages".D011.Rows[11].Used OR "FRK_PersistImages".D011.Rows[11].SchemaVersion <> 4 OR "FRK_PersistImages".D011.Rows[11].ModelCode <> 'MODEL_B' OR "FRK_PersistImages".D011.Rows[11].Record.Scope <> 'StationB.Satellite.Cell' OR "FRK_PersistImages".D011.Rows[11].Record.WriteKey <> 'timeout' OR "FRK_PersistImages".D011.Rows[11].Record.Revision <> 1 OR "FRK_PersistImages".D011.Rows[11].Record.Kind <> 0 OR "FRK_PersistImages".D011.Rows[11].Record.ValueType <> 3 THEN RETURN; END_IF;
    #Ok := "FRK_ConfigDecode"(Text := STRING_TO_WSTRING("FRK_PersistImages".D011.Rows[11].Record.ValueText), Storage := 7, Minimum := 1.0, Maximum := 60000.0, MaxLength := 0, Value := "FRK_ConfigScratch".Value);
    IF NOT #Ok THEN RETURN; END_IF;
    IF NOT "FRK_PersistImages".D011.Rows[12].Used OR "FRK_PersistImages".D011.Rows[12].SchemaVersion <> 4 OR "FRK_PersistImages".D011.Rows[12].ModelCode <> 'MODEL_B' OR "FRK_PersistImages".D011.Rows[12].Record.Scope <> 'StationB.Satellite.Cell' OR "FRK_PersistImages".D011.Rows[12].Record.WriteKey <> 'preset' OR "FRK_PersistImages".D011.Rows[12].Record.Revision <> 2 OR "FRK_PersistImages".D011.Rows[12].Record.Kind <> 0 OR "FRK_PersistImages".D011.Rows[12].Record.ValueType <> 0 THEN RETURN; END_IF;
    #Ok := "FRK_ConfigDecode"(Text := STRING_TO_WSTRING("FRK_PersistImages".D011.Rows[12].Record.ValueText), Storage := 3, Minimum := 0.0, Maximum := 1000.0, MaxLength := 0, Value := "FRK_ConfigScratch".Value);
    IF NOT #Ok THEN RETURN; END_IF;
    IF NOT "FRK_PersistImages".D011.Rows[13].Used OR "FRK_PersistImages".D011.Rows[13].SchemaVersion <> 4 OR "FRK_PersistImages".D011.Rows[13].ModelCode <> 'MODEL_B' OR "FRK_PersistImages".D011.Rows[13].Record.Scope <> 'StationB.Satellite.Cell.Clamp' OR "FRK_PersistImages".D011.Rows[13].Record.WriteKey <> 'timeout' OR "FRK_PersistImages".D011.Rows[13].Record.Revision <> 1 OR "FRK_PersistImages".D011.Rows[13].Record.Kind <> 0 OR "FRK_PersistImages".D011.Rows[13].Record.ValueType <> 3 THEN RETURN; END_IF;
    #Ok := "FRK_ConfigDecode"(Text := STRING_TO_WSTRING("FRK_PersistImages".D011.Rows[13].Record.ValueText), Storage := 7, Minimum := 1.0, Maximum := 60000.0, MaxLength := 0, Value := "FRK_ConfigScratch".Value);
    IF NOT #Ok THEN RETURN; END_IF;
    IF NOT "FRK_PersistImages".D011.Rows[14].Used OR "FRK_PersistImages".D011.Rows[14].SchemaVersion <> 4 OR "FRK_PersistImages".D011.Rows[14].ModelCode <> 'MODEL_B' OR "FRK_PersistImages".D011.Rows[14].Record.Scope <> 'StationB.Satellite.Cell.Clamp' OR "FRK_PersistImages".D011.Rows[14].Record.WriteKey <> 'preset' OR "FRK_PersistImages".D011.Rows[14].Record.Revision <> 2 OR "FRK_PersistImages".D011.Rows[14].Record.Kind <> 0 OR "FRK_PersistImages".D011.Rows[14].Record.ValueType <> 0 THEN RETURN; END_IF;
    #Ok := "FRK_ConfigDecode"(Text := STRING_TO_WSTRING("FRK_PersistImages".D011.Rows[14].Record.ValueText), Storage := 3, Minimum := 0.0, Maximum := 1000.0, MaxLength := 0, Value := "FRK_ConfigScratch".Value);
    IF NOT #Ok THEN RETURN; END_IF;
    IF NOT "FRK_PersistImages".D011.Rows[15].Used OR "FRK_PersistImages".D011.Rows[15].SchemaVersion <> 4 OR "FRK_PersistImages".D011.Rows[15].ModelCode <> 'MODEL_B' OR "FRK_PersistImages".D011.Rows[15].Record.Scope <> 'StationB.Satellite.Cell.Gate' OR "FRK_PersistImages".D011.Rows[15].Record.WriteKey <> 'timeout' OR "FRK_PersistImages".D011.Rows[15].Record.Revision <> 1 OR "FRK_PersistImages".D011.Rows[15].Record.Kind <> 0 OR "FRK_PersistImages".D011.Rows[15].Record.ValueType <> 3 THEN RETURN; END_IF;
    #Ok := "FRK_ConfigDecode"(Text := STRING_TO_WSTRING("FRK_PersistImages".D011.Rows[15].Record.ValueText), Storage := 7, Minimum := 1.0, Maximum := 60000.0, MaxLength := 0, Value := "FRK_ConfigScratch".Value);
    IF NOT #Ok THEN RETURN; END_IF;
    IF NOT "FRK_PersistImages".D011.Rows[16].Used OR "FRK_PersistImages".D011.Rows[16].SchemaVersion <> 4 OR "FRK_PersistImages".D011.Rows[16].ModelCode <> 'MODEL_B' OR "FRK_PersistImages".D011.Rows[16].Record.Scope <> 'StationB.Satellite.Cell.Gate' OR "FRK_PersistImages".D011.Rows[16].Record.WriteKey <> 'preset' OR "FRK_PersistImages".D011.Rows[16].Record.Revision <> 2 OR "FRK_PersistImages".D011.Rows[16].Record.Kind <> 0 OR "FRK_PersistImages".D011.Rows[16].Record.ValueType <> 0 THEN RETURN; END_IF;
    #Ok := "FRK_ConfigDecode"(Text := STRING_TO_WSTRING("FRK_PersistImages".D011.Rows[16].Record.ValueText), Storage := 3, Minimum := 0.0, Maximum := 1000.0, MaxLength := 0, Value := "FRK_ConfigScratch".Value);
    IF NOT #Ok THEN RETURN; END_IF;
    IF NOT "FRK_PersistImages".D011.Rows[17].Used OR "FRK_PersistImages".D011.Rows[17].SchemaVersion <> 4 OR "FRK_PersistImages".D011.Rows[17].ModelCode <> 'MODEL_B' OR "FRK_PersistImages".D011.Rows[17].Record.Scope <> 'StationB.Satellite.Inner' OR "FRK_PersistImages".D011.Rows[17].Record.WriteKey <> 'timeout' OR "FRK_PersistImages".D011.Rows[17].Record.Revision <> 1 OR "FRK_PersistImages".D011.Rows[17].Record.Kind <> 0 OR "FRK_PersistImages".D011.Rows[17].Record.ValueType <> 3 THEN RETURN; END_IF;
    #Ok := "FRK_ConfigDecode"(Text := STRING_TO_WSTRING("FRK_PersistImages".D011.Rows[17].Record.ValueText), Storage := 7, Minimum := 1.0, Maximum := 60000.0, MaxLength := 0, Value := "FRK_ConfigScratch".Value);
    IF NOT #Ok THEN RETURN; END_IF;
    IF NOT "FRK_PersistImages".D011.Rows[18].Used OR "FRK_PersistImages".D011.Rows[18].SchemaVersion <> 4 OR "FRK_PersistImages".D011.Rows[18].ModelCode <> 'MODEL_B' OR "FRK_PersistImages".D011.Rows[18].Record.Scope <> 'StationB.Satellite.Inner' OR "FRK_PersistImages".D011.Rows[18].Record.WriteKey <> 'preset' OR "FRK_PersistImages".D011.Rows[18].Record.Revision <> 2 OR "FRK_PersistImages".D011.Rows[18].Record.Kind <> 0 OR "FRK_PersistImages".D011.Rows[18].Record.ValueType <> 0 THEN RETURN; END_IF;
    #Ok := "FRK_ConfigDecode"(Text := STRING_TO_WSTRING("FRK_PersistImages".D011.Rows[18].Record.ValueText), Storage := 3, Minimum := 0.0, Maximum := 1000.0, MaxLength := 0, Value := "FRK_ConfigScratch".Value);
    IF NOT #Ok THEN RETURN; END_IF;
    IF NOT "FRK_PersistImages".D011.Rows[19].Used OR "FRK_PersistImages".D011.Rows[19].SchemaVersion <> 4 OR "FRK_PersistImages".D011.Rows[19].ModelCode <> 'MODEL_B' OR "FRK_PersistImages".D011.Rows[19].Record.Scope <> 'StationB.Satellite.Inner.Cell' OR "FRK_PersistImages".D011.Rows[19].Record.WriteKey <> 'timeout' OR "FRK_PersistImages".D011.Rows[19].Record.Revision <> 1 OR "FRK_PersistImages".D011.Rows[19].Record.Kind <> 0 OR "FRK_PersistImages".D011.Rows[19].Record.ValueType <> 3 THEN RETURN; END_IF;
    #Ok := "FRK_ConfigDecode"(Text := STRING_TO_WSTRING("FRK_PersistImages".D011.Rows[19].Record.ValueText), Storage := 7, Minimum := 1.0, Maximum := 60000.0, MaxLength := 0, Value := "FRK_ConfigScratch".Value);
    IF NOT #Ok THEN RETURN; END_IF;
    IF NOT "FRK_PersistImages".D011.Rows[20].Used OR "FRK_PersistImages".D011.Rows[20].SchemaVersion <> 4 OR "FRK_PersistImages".D011.Rows[20].ModelCode <> 'MODEL_B' OR "FRK_PersistImages".D011.Rows[20].Record.Scope <> 'StationB.Satellite.Inner.Cell' OR "FRK_PersistImages".D011.Rows[20].Record.WriteKey <> 'preset' OR "FRK_PersistImages".D011.Rows[20].Record.Revision <> 2 OR "FRK_PersistImages".D011.Rows[20].Record.Kind <> 0 OR "FRK_PersistImages".D011.Rows[20].Record.ValueType <> 0 THEN RETURN; END_IF;
    #Ok := "FRK_ConfigDecode"(Text := STRING_TO_WSTRING("FRK_PersistImages".D011.Rows[20].Record.ValueText), Storage := 3, Minimum := 0.0, Maximum := 1000.0, MaxLength := 0, Value := "FRK_ConfigScratch".Value);
    IF NOT #Ok THEN RETURN; END_IF;
    IF NOT "FRK_PersistImages".D011.Rows[21].Used OR "FRK_PersistImages".D011.Rows[21].SchemaVersion <> 4 OR "FRK_PersistImages".D011.Rows[21].ModelCode <> 'MODEL_B' OR "FRK_PersistImages".D011.Rows[21].Record.Scope <> 'StationB.Satellite.Inner.Cell.Clamp' OR "FRK_PersistImages".D011.Rows[21].Record.WriteKey <> 'timeout' OR "FRK_PersistImages".D011.Rows[21].Record.Revision <> 1 OR "FRK_PersistImages".D011.Rows[21].Record.Kind <> 0 OR "FRK_PersistImages".D011.Rows[21].Record.ValueType <> 3 THEN RETURN; END_IF;
    #Ok := "FRK_ConfigDecode"(Text := STRING_TO_WSTRING("FRK_PersistImages".D011.Rows[21].Record.ValueText), Storage := 7, Minimum := 1.0, Maximum := 60000.0, MaxLength := 0, Value := "FRK_ConfigScratch".Value);
    IF NOT #Ok THEN RETURN; END_IF;
    IF NOT "FRK_PersistImages".D011.Rows[22].Used OR "FRK_PersistImages".D011.Rows[22].SchemaVersion <> 4 OR "FRK_PersistImages".D011.Rows[22].ModelCode <> 'MODEL_B' OR "FRK_PersistImages".D011.Rows[22].Record.Scope <> 'StationB.Satellite.Inner.Cell.Clamp' OR "FRK_PersistImages".D011.Rows[22].Record.WriteKey <> 'preset' OR "FRK_PersistImages".D011.Rows[22].Record.Revision <> 2 OR "FRK_PersistImages".D011.Rows[22].Record.Kind <> 0 OR "FRK_PersistImages".D011.Rows[22].Record.ValueType <> 0 THEN RETURN; END_IF;
    #Ok := "FRK_ConfigDecode"(Text := STRING_TO_WSTRING("FRK_PersistImages".D011.Rows[22].Record.ValueText), Storage := 3, Minimum := 0.0, Maximum := 1000.0, MaxLength := 0, Value := "FRK_ConfigScratch".Value);
    IF NOT #Ok THEN RETURN; END_IF;
    IF NOT "FRK_PersistImages".D011.Rows[23].Used OR "FRK_PersistImages".D011.Rows[23].SchemaVersion <> 4 OR "FRK_PersistImages".D011.Rows[23].ModelCode <> 'MODEL_B' OR "FRK_PersistImages".D011.Rows[23].Record.Scope <> 'StationB.Satellite.Inner.Cell.Gate' OR "FRK_PersistImages".D011.Rows[23].Record.WriteKey <> 'timeout' OR "FRK_PersistImages".D011.Rows[23].Record.Revision <> 1 OR "FRK_PersistImages".D011.Rows[23].Record.Kind <> 0 OR "FRK_PersistImages".D011.Rows[23].Record.ValueType <> 3 THEN RETURN; END_IF;
    #Ok := "FRK_ConfigDecode"(Text := STRING_TO_WSTRING("FRK_PersistImages".D011.Rows[23].Record.ValueText), Storage := 7, Minimum := 1.0, Maximum := 60000.0, MaxLength := 0, Value := "FRK_ConfigScratch".Value);
    IF NOT #Ok THEN RETURN; END_IF;
    IF NOT "FRK_PersistImages".D011.Rows[24].Used OR "FRK_PersistImages".D011.Rows[24].SchemaVersion <> 4 OR "FRK_PersistImages".D011.Rows[24].ModelCode <> 'MODEL_B' OR "FRK_PersistImages".D011.Rows[24].Record.Scope <> 'StationB.Satellite.Inner.Cell.Gate' OR "FRK_PersistImages".D011.Rows[24].Record.WriteKey <> 'preset' OR "FRK_PersistImages".D011.Rows[24].Record.Revision <> 2 OR "FRK_PersistImages".D011.Rows[24].Record.Kind <> 0 OR "FRK_PersistImages".D011.Rows[24].Record.ValueType <> 0 THEN RETURN; END_IF;
    #Ok := "FRK_ConfigDecode"(Text := STRING_TO_WSTRING("FRK_PersistImages".D011.Rows[24].Record.ValueText), Storage := 3, Minimum := 0.0, Maximum := 1000.0, MaxLength := 0, Value := "FRK_ConfigScratch".Value);
    IF NOT #Ok THEN RETURN; END_IF;
    #Stored := "FRK_ConfigFind"(Scope := 'StationB', Key := 'timeout', ModelCode := 'MODEL_B');
    IF #Stored = 0 THEN
        FOR #Index := 1 TO 114 DO
            #Reserved := NOT "FRK_ConfigStore".Rows[#Index].Used;
            FOR #Prior := 1 TO 0 DO IF #Targets[#Prior] = #Index THEN #Reserved := FALSE; END_IF; END_FOR;
            IF #Reserved THEN #Stored := #Index; EXIT; END_IF;
        END_FOR;
    END_IF;
    IF #Stored < 1 OR #Stored > 114 THEN RETURN; END_IF;
    #Targets[1] := #Stored;
    #Stored := "FRK_ConfigFind"(Scope := 'StationB', Key := 'preset', ModelCode := 'MODEL_B');
    IF #Stored = 0 THEN
        FOR #Index := 1 TO 114 DO
            #Reserved := NOT "FRK_ConfigStore".Rows[#Index].Used;
            FOR #Prior := 1 TO 1 DO IF #Targets[#Prior] = #Index THEN #Reserved := FALSE; END_IF; END_FOR;
            IF #Reserved THEN #Stored := #Index; EXIT; END_IF;
        END_FOR;
    END_IF;
    IF #Stored < 1 OR #Stored > 114 THEN RETURN; END_IF;
    #Targets[2] := #Stored;
    #Stored := "FRK_ConfigFind"(Scope := 'StationB.Cell', Key := 'timeout', ModelCode := 'MODEL_B');
    IF #Stored = 0 THEN
        FOR #Index := 1 TO 114 DO
            #Reserved := NOT "FRK_ConfigStore".Rows[#Index].Used;
            FOR #Prior := 1 TO 2 DO IF #Targets[#Prior] = #Index THEN #Reserved := FALSE; END_IF; END_FOR;
            IF #Reserved THEN #Stored := #Index; EXIT; END_IF;
        END_FOR;
    END_IF;
    IF #Stored < 1 OR #Stored > 114 THEN RETURN; END_IF;
    #Targets[3] := #Stored;
    #Stored := "FRK_ConfigFind"(Scope := 'StationB.Cell', Key := 'preset', ModelCode := 'MODEL_B');
    IF #Stored = 0 THEN
        FOR #Index := 1 TO 114 DO
            #Reserved := NOT "FRK_ConfigStore".Rows[#Index].Used;
            FOR #Prior := 1 TO 3 DO IF #Targets[#Prior] = #Index THEN #Reserved := FALSE; END_IF; END_FOR;
            IF #Reserved THEN #Stored := #Index; EXIT; END_IF;
        END_FOR;
    END_IF;
    IF #Stored < 1 OR #Stored > 114 THEN RETURN; END_IF;
    #Targets[4] := #Stored;
    #Stored := "FRK_ConfigFind"(Scope := 'StationB.Cell.Clamp', Key := 'timeout', ModelCode := 'MODEL_B');
    IF #Stored = 0 THEN
        FOR #Index := 1 TO 114 DO
            #Reserved := NOT "FRK_ConfigStore".Rows[#Index].Used;
            FOR #Prior := 1 TO 4 DO IF #Targets[#Prior] = #Index THEN #Reserved := FALSE; END_IF; END_FOR;
            IF #Reserved THEN #Stored := #Index; EXIT; END_IF;
        END_FOR;
    END_IF;
    IF #Stored < 1 OR #Stored > 114 THEN RETURN; END_IF;
    #Targets[5] := #Stored;
    #Stored := "FRK_ConfigFind"(Scope := 'StationB.Cell.Clamp', Key := 'preset', ModelCode := 'MODEL_B');
    IF #Stored = 0 THEN
        FOR #Index := 1 TO 114 DO
            #Reserved := NOT "FRK_ConfigStore".Rows[#Index].Used;
            FOR #Prior := 1 TO 5 DO IF #Targets[#Prior] = #Index THEN #Reserved := FALSE; END_IF; END_FOR;
            IF #Reserved THEN #Stored := #Index; EXIT; END_IF;
        END_FOR;
    END_IF;
    IF #Stored < 1 OR #Stored > 114 THEN RETURN; END_IF;
    #Targets[6] := #Stored;
    #Stored := "FRK_ConfigFind"(Scope := 'StationB.Cell.Gate', Key := 'timeout', ModelCode := 'MODEL_B');
    IF #Stored = 0 THEN
        FOR #Index := 1 TO 114 DO
            #Reserved := NOT "FRK_ConfigStore".Rows[#Index].Used;
            FOR #Prior := 1 TO 6 DO IF #Targets[#Prior] = #Index THEN #Reserved := FALSE; END_IF; END_FOR;
            IF #Reserved THEN #Stored := #Index; EXIT; END_IF;
        END_FOR;
    END_IF;
    IF #Stored < 1 OR #Stored > 114 THEN RETURN; END_IF;
    #Targets[7] := #Stored;
    #Stored := "FRK_ConfigFind"(Scope := 'StationB.Cell.Gate', Key := 'preset', ModelCode := 'MODEL_B');
    IF #Stored = 0 THEN
        FOR #Index := 1 TO 114 DO
            #Reserved := NOT "FRK_ConfigStore".Rows[#Index].Used;
            FOR #Prior := 1 TO 7 DO IF #Targets[#Prior] = #Index THEN #Reserved := FALSE; END_IF; END_FOR;
            IF #Reserved THEN #Stored := #Index; EXIT; END_IF;
        END_FOR;
    END_IF;
    IF #Stored < 1 OR #Stored > 114 THEN RETURN; END_IF;
    #Targets[8] := #Stored;
    #Stored := "FRK_ConfigFind"(Scope := 'StationB.Satellite', Key := 'timeout', ModelCode := 'MODEL_B');
    IF #Stored = 0 THEN
        FOR #Index := 1 TO 114 DO
            #Reserved := NOT "FRK_ConfigStore".Rows[#Index].Used;
            FOR #Prior := 1 TO 8 DO IF #Targets[#Prior] = #Index THEN #Reserved := FALSE; END_IF; END_FOR;
            IF #Reserved THEN #Stored := #Index; EXIT; END_IF;
        END_FOR;
    END_IF;
    IF #Stored < 1 OR #Stored > 114 THEN RETURN; END_IF;
    #Targets[9] := #Stored;
    #Stored := "FRK_ConfigFind"(Scope := 'StationB.Satellite', Key := 'preset', ModelCode := 'MODEL_B');
    IF #Stored = 0 THEN
        FOR #Index := 1 TO 114 DO
            #Reserved := NOT "FRK_ConfigStore".Rows[#Index].Used;
            FOR #Prior := 1 TO 9 DO IF #Targets[#Prior] = #Index THEN #Reserved := FALSE; END_IF; END_FOR;
            IF #Reserved THEN #Stored := #Index; EXIT; END_IF;
        END_FOR;
    END_IF;
    IF #Stored < 1 OR #Stored > 114 THEN RETURN; END_IF;
    #Targets[10] := #Stored;
    #Stored := "FRK_ConfigFind"(Scope := 'StationB.Satellite.Cell', Key := 'timeout', ModelCode := 'MODEL_B');
    IF #Stored = 0 THEN
        FOR #Index := 1 TO 114 DO
            #Reserved := NOT "FRK_ConfigStore".Rows[#Index].Used;
            FOR #Prior := 1 TO 10 DO IF #Targets[#Prior] = #Index THEN #Reserved := FALSE; END_IF; END_FOR;
            IF #Reserved THEN #Stored := #Index; EXIT; END_IF;
        END_FOR;
    END_IF;
    IF #Stored < 1 OR #Stored > 114 THEN RETURN; END_IF;
    #Targets[11] := #Stored;
    #Stored := "FRK_ConfigFind"(Scope := 'StationB.Satellite.Cell', Key := 'preset', ModelCode := 'MODEL_B');
    IF #Stored = 0 THEN
        FOR #Index := 1 TO 114 DO
            #Reserved := NOT "FRK_ConfigStore".Rows[#Index].Used;
            FOR #Prior := 1 TO 11 DO IF #Targets[#Prior] = #Index THEN #Reserved := FALSE; END_IF; END_FOR;
            IF #Reserved THEN #Stored := #Index; EXIT; END_IF;
        END_FOR;
    END_IF;
    IF #Stored < 1 OR #Stored > 114 THEN RETURN; END_IF;
    #Targets[12] := #Stored;
    #Stored := "FRK_ConfigFind"(Scope := 'StationB.Satellite.Cell.Clamp', Key := 'timeout', ModelCode := 'MODEL_B');
    IF #Stored = 0 THEN
        FOR #Index := 1 TO 114 DO
            #Reserved := NOT "FRK_ConfigStore".Rows[#Index].Used;
            FOR #Prior := 1 TO 12 DO IF #Targets[#Prior] = #Index THEN #Reserved := FALSE; END_IF; END_FOR;
            IF #Reserved THEN #Stored := #Index; EXIT; END_IF;
        END_FOR;
    END_IF;
    IF #Stored < 1 OR #Stored > 114 THEN RETURN; END_IF;
    #Targets[13] := #Stored;
    #Stored := "FRK_ConfigFind"(Scope := 'StationB.Satellite.Cell.Clamp', Key := 'preset', ModelCode := 'MODEL_B');
    IF #Stored = 0 THEN
        FOR #Index := 1 TO 114 DO
            #Reserved := NOT "FRK_ConfigStore".Rows[#Index].Used;
            FOR #Prior := 1 TO 13 DO IF #Targets[#Prior] = #Index THEN #Reserved := FALSE; END_IF; END_FOR;
            IF #Reserved THEN #Stored := #Index; EXIT; END_IF;
        END_FOR;
    END_IF;
    IF #Stored < 1 OR #Stored > 114 THEN RETURN; END_IF;
    #Targets[14] := #Stored;
    #Stored := "FRK_ConfigFind"(Scope := 'StationB.Satellite.Cell.Gate', Key := 'timeout', ModelCode := 'MODEL_B');
    IF #Stored = 0 THEN
        FOR #Index := 1 TO 114 DO
            #Reserved := NOT "FRK_ConfigStore".Rows[#Index].Used;
            FOR #Prior := 1 TO 14 DO IF #Targets[#Prior] = #Index THEN #Reserved := FALSE; END_IF; END_FOR;
            IF #Reserved THEN #Stored := #Index; EXIT; END_IF;
        END_FOR;
    END_IF;
    IF #Stored < 1 OR #Stored > 114 THEN RETURN; END_IF;
    #Targets[15] := #Stored;
    #Stored := "FRK_ConfigFind"(Scope := 'StationB.Satellite.Cell.Gate', Key := 'preset', ModelCode := 'MODEL_B');
    IF #Stored = 0 THEN
        FOR #Index := 1 TO 114 DO
            #Reserved := NOT "FRK_ConfigStore".Rows[#Index].Used;
            FOR #Prior := 1 TO 15 DO IF #Targets[#Prior] = #Index THEN #Reserved := FALSE; END_IF; END_FOR;
            IF #Reserved THEN #Stored := #Index; EXIT; END_IF;
        END_FOR;
    END_IF;
    IF #Stored < 1 OR #Stored > 114 THEN RETURN; END_IF;
    #Targets[16] := #Stored;
    #Stored := "FRK_ConfigFind"(Scope := 'StationB.Satellite.Inner', Key := 'timeout', ModelCode := 'MODEL_B');
    IF #Stored = 0 THEN
        FOR #Index := 1 TO 114 DO
            #Reserved := NOT "FRK_ConfigStore".Rows[#Index].Used;
            FOR #Prior := 1 TO 16 DO IF #Targets[#Prior] = #Index THEN #Reserved := FALSE; END_IF; END_FOR;
            IF #Reserved THEN #Stored := #Index; EXIT; END_IF;
        END_FOR;
    END_IF;
    IF #Stored < 1 OR #Stored > 114 THEN RETURN; END_IF;
    #Targets[17] := #Stored;
    #Stored := "FRK_ConfigFind"(Scope := 'StationB.Satellite.Inner', Key := 'preset', ModelCode := 'MODEL_B');
    IF #Stored = 0 THEN
        FOR #Index := 1 TO 114 DO
            #Reserved := NOT "FRK_ConfigStore".Rows[#Index].Used;
            FOR #Prior := 1 TO 17 DO IF #Targets[#Prior] = #Index THEN #Reserved := FALSE; END_IF; END_FOR;
            IF #Reserved THEN #Stored := #Index; EXIT; END_IF;
        END_FOR;
    END_IF;
    IF #Stored < 1 OR #Stored > 114 THEN RETURN; END_IF;
    #Targets[18] := #Stored;
    #Stored := "FRK_ConfigFind"(Scope := 'StationB.Satellite.Inner.Cell', Key := 'timeout', ModelCode := 'MODEL_B');
    IF #Stored = 0 THEN
        FOR #Index := 1 TO 114 DO
            #Reserved := NOT "FRK_ConfigStore".Rows[#Index].Used;
            FOR #Prior := 1 TO 18 DO IF #Targets[#Prior] = #Index THEN #Reserved := FALSE; END_IF; END_FOR;
            IF #Reserved THEN #Stored := #Index; EXIT; END_IF;
        END_FOR;
    END_IF;
    IF #Stored < 1 OR #Stored > 114 THEN RETURN; END_IF;
    #Targets[19] := #Stored;
    #Stored := "FRK_ConfigFind"(Scope := 'StationB.Satellite.Inner.Cell', Key := 'preset', ModelCode := 'MODEL_B');
    IF #Stored = 0 THEN
        FOR #Index := 1 TO 114 DO
            #Reserved := NOT "FRK_ConfigStore".Rows[#Index].Used;
            FOR #Prior := 1 TO 19 DO IF #Targets[#Prior] = #Index THEN #Reserved := FALSE; END_IF; END_FOR;
            IF #Reserved THEN #Stored := #Index; EXIT; END_IF;
        END_FOR;
    END_IF;
    IF #Stored < 1 OR #Stored > 114 THEN RETURN; END_IF;
    #Targets[20] := #Stored;
    #Stored := "FRK_ConfigFind"(Scope := 'StationB.Satellite.Inner.Cell.Clamp', Key := 'timeout', ModelCode := 'MODEL_B');
    IF #Stored = 0 THEN
        FOR #Index := 1 TO 114 DO
            #Reserved := NOT "FRK_ConfigStore".Rows[#Index].Used;
            FOR #Prior := 1 TO 20 DO IF #Targets[#Prior] = #Index THEN #Reserved := FALSE; END_IF; END_FOR;
            IF #Reserved THEN #Stored := #Index; EXIT; END_IF;
        END_FOR;
    END_IF;
    IF #Stored < 1 OR #Stored > 114 THEN RETURN; END_IF;
    #Targets[21] := #Stored;
    #Stored := "FRK_ConfigFind"(Scope := 'StationB.Satellite.Inner.Cell.Clamp', Key := 'preset', ModelCode := 'MODEL_B');
    IF #Stored = 0 THEN
        FOR #Index := 1 TO 114 DO
            #Reserved := NOT "FRK_ConfigStore".Rows[#Index].Used;
            FOR #Prior := 1 TO 21 DO IF #Targets[#Prior] = #Index THEN #Reserved := FALSE; END_IF; END_FOR;
            IF #Reserved THEN #Stored := #Index; EXIT; END_IF;
        END_FOR;
    END_IF;
    IF #Stored < 1 OR #Stored > 114 THEN RETURN; END_IF;
    #Targets[22] := #Stored;
    #Stored := "FRK_ConfigFind"(Scope := 'StationB.Satellite.Inner.Cell.Gate', Key := 'timeout', ModelCode := 'MODEL_B');
    IF #Stored = 0 THEN
        FOR #Index := 1 TO 114 DO
            #Reserved := NOT "FRK_ConfigStore".Rows[#Index].Used;
            FOR #Prior := 1 TO 22 DO IF #Targets[#Prior] = #Index THEN #Reserved := FALSE; END_IF; END_FOR;
            IF #Reserved THEN #Stored := #Index; EXIT; END_IF;
        END_FOR;
    END_IF;
    IF #Stored < 1 OR #Stored > 114 THEN RETURN; END_IF;
    #Targets[23] := #Stored;
    #Stored := "FRK_ConfigFind"(Scope := 'StationB.Satellite.Inner.Cell.Gate', Key := 'preset', ModelCode := 'MODEL_B');
    IF #Stored = 0 THEN
        FOR #Index := 1 TO 114 DO
            #Reserved := NOT "FRK_ConfigStore".Rows[#Index].Used;
            FOR #Prior := 1 TO 23 DO IF #Targets[#Prior] = #Index THEN #Reserved := FALSE; END_IF; END_FOR;
            IF #Reserved THEN #Stored := #Index; EXIT; END_IF;
        END_FOR;
    END_IF;
    IF #Stored < 1 OR #Stored > 114 THEN RETURN; END_IF;
    #Targets[24] := #Stored;
    "FRK_ConfigStore".Rows[#Targets[1]] := "FRK_PersistImages".D011.Rows[1];
    "FRK_ConfigStore".Rows[#Targets[2]] := "FRK_PersistImages".D011.Rows[2];
    "FRK_ConfigStore".Rows[#Targets[3]] := "FRK_PersistImages".D011.Rows[3];
    "FRK_ConfigStore".Rows[#Targets[4]] := "FRK_PersistImages".D011.Rows[4];
    "FRK_ConfigStore".Rows[#Targets[5]] := "FRK_PersistImages".D011.Rows[5];
    "FRK_ConfigStore".Rows[#Targets[6]] := "FRK_PersistImages".D011.Rows[6];
    "FRK_ConfigStore".Rows[#Targets[7]] := "FRK_PersistImages".D011.Rows[7];
    "FRK_ConfigStore".Rows[#Targets[8]] := "FRK_PersistImages".D011.Rows[8];
    "FRK_ConfigStore".Rows[#Targets[9]] := "FRK_PersistImages".D011.Rows[9];
    "FRK_ConfigStore".Rows[#Targets[10]] := "FRK_PersistImages".D011.Rows[10];
    "FRK_ConfigStore".Rows[#Targets[11]] := "FRK_PersistImages".D011.Rows[11];
    "FRK_ConfigStore".Rows[#Targets[12]] := "FRK_PersistImages".D011.Rows[12];
    "FRK_ConfigStore".Rows[#Targets[13]] := "FRK_PersistImages".D011.Rows[13];
    "FRK_ConfigStore".Rows[#Targets[14]] := "FRK_PersistImages".D011.Rows[14];
    "FRK_ConfigStore".Rows[#Targets[15]] := "FRK_PersistImages".D011.Rows[15];
    "FRK_ConfigStore".Rows[#Targets[16]] := "FRK_PersistImages".D011.Rows[16];
    "FRK_ConfigStore".Rows[#Targets[17]] := "FRK_PersistImages".D011.Rows[17];
    "FRK_ConfigStore".Rows[#Targets[18]] := "FRK_PersistImages".D011.Rows[18];
    "FRK_ConfigStore".Rows[#Targets[19]] := "FRK_PersistImages".D011.Rows[19];
    "FRK_ConfigStore".Rows[#Targets[20]] := "FRK_PersistImages".D011.Rows[20];
    "FRK_ConfigStore".Rows[#Targets[21]] := "FRK_PersistImages".D011.Rows[21];
    "FRK_ConfigStore".Rows[#Targets[22]] := "FRK_PersistImages".D011.Rows[22];
    "FRK_ConfigStore".Rows[#Targets[23]] := "FRK_PersistImages".D011.Rows[23];
    "FRK_ConfigStore".Rows[#Targets[24]] := "FRK_PersistImages".D011.Rows[24];
    "FRK_ConfigStore".SchemaVersion := 1;
    #FRK_DocApply_D011 := TRUE;
END_FUNCTION
FUNCTION "FRK_DocCapture_D012" : Bool
{ S7_Optimized_Access := 'TRUE' }
VERSION : 0.1
VAR_IN_OUT
    Length : DInt;
END_VAR
VAR_TEMP
    Index : Int;
    Stored : Int;
    Position : DInt;
    NativeResult : Int;
    Ok : Bool;
END_VAR
BEGIN
    #FRK_DocCapture_D012 := FALSE;
    "FRK_PersistImages".D012.SchemaVersion := 1; "FRK_PersistImages".D012.Scope := 'StationB';
    #Stored := 0;
    FOR #Index := 1 TO 2 DO
        IF "FRK_AccessPolicies".Rows[#Index].Scope = 'StationB' THEN #Stored := #Index; END_IF;
    END_FOR;
    IF #Stored = 0 THEN RETURN; END_IF;
    "FRK_PersistImages".D012.Image := "FRK_AccessPolicies".Rows[#Stored];
    IF NOT "FRK_AccessPolicyValid"(Image := "FRK_PersistImages".D012.Image) THEN RETURN; END_IF;
    FOR #Index := 0 TO 413 DO "FRK_PersistBuffers".D012Data[#Index] := BYTE#0; END_FOR;
    #Position := 24;
    #NativeResult := Serialize(SRC_VARIABLE := "FRK_PersistImages".D012, DEST_ARRAY => "FRK_PersistBuffers".D012Data, POS := #Position);
    IF #NativeResult <> 0 OR #Position < 24 OR #Position > 414 THEN RETURN; END_IF;
    #Length := #Position - 24;
    #FRK_DocCapture_D012 := TRUE;
END_FUNCTION
FUNCTION "FRK_DocApply_D012" : Bool
{ S7_Optimized_Access := 'TRUE' }
VERSION : 0.1
VAR_TEMP
    Index : Int;
    Stored : Int;
    Position : DInt;
    NativeResult : Int;
    Ok : Bool;
END_VAR
BEGIN
    #FRK_DocApply_D012 := FALSE;
    #Position := 24;
    #NativeResult := Deserialize(SRC_ARRAY := "FRK_PersistBuffers".D012Data, DEST_VARIABLE => "FRK_PersistImages".D012, POS := #Position);
    IF #NativeResult <> 0 OR #Position <> 24 + UDINT_TO_DINT("FRK_PersistConsumers".Rows[12].Result.Length) THEN RETURN; END_IF;
    IF "FRK_PersistImages".D012.SchemaVersion <> 1 OR "FRK_PersistImages".D012.Scope <> 'StationB' THEN RETURN; END_IF;
    IF "FRK_PersistImages".D012.Image.Scope <> 'StationB' OR NOT "FRK_AccessPolicyValid"(Image := "FRK_PersistImages".D012.Image) THEN RETURN; END_IF;
    "FRK_AccessPolicies".Rows[2] := "FRK_PersistImages".D012.Image;
    #FRK_DocApply_D012 := TRUE;
END_FUNCTION
FUNCTION "FRK_DocCapture_D013" : Bool
{ S7_Optimized_Access := 'TRUE' }
VERSION : 0.1
VAR_IN_OUT
    Length : DInt;
END_VAR
VAR_TEMP
    Index : Int;
    Stored : Int;
    Position : DInt;
    NativeResult : Int;
    Ok : Bool;
END_VAR
BEGIN
    #FRK_DocCapture_D013 := FALSE;
    "FRK_PersistImages".D013.SchemaVersion := 1; "FRK_PersistImages".D013.Scope := 'StationB';
    "FRK_PersistImages".D013.Ordinal := 1;
    "FRK_PersistImages".D013.Payload := "FRK_SetStore".Sets[2, 1];
    FOR #Index := 0 TO 9359 DO "FRK_PersistBuffers".D013Data[#Index] := BYTE#0; END_FOR;
    #Position := 24;
    #NativeResult := Serialize(SRC_VARIABLE := "FRK_PersistImages".D013, DEST_ARRAY => "FRK_PersistBuffers".D013Data, POS := #Position);
    IF #NativeResult <> 0 OR #Position < 24 OR #Position > 9360 THEN RETURN; END_IF;
    #Length := #Position - 24;
    #FRK_DocCapture_D013 := TRUE;
END_FUNCTION
FUNCTION "FRK_DocApply_D013" : Bool
{ S7_Optimized_Access := 'TRUE' }
VERSION : 0.1
VAR_TEMP
    Index : Int;
    Stored : Int;
    Position : DInt;
    NativeResult : Int;
    Ok : Bool;
END_VAR
BEGIN
    #FRK_DocApply_D013 := FALSE;
    #Position := 24;
    #NativeResult := Deserialize(SRC_ARRAY := "FRK_PersistBuffers".D013Data, DEST_VARIABLE => "FRK_PersistImages".D013, POS := #Position);
    IF #NativeResult <> 0 OR #Position <> 24 + UDINT_TO_DINT("FRK_PersistConsumers".Rows[13].Result.Length) THEN RETURN; END_IF;
    IF "FRK_PersistImages".D013.SchemaVersion <> 1 OR "FRK_PersistImages".D013.Scope <> 'StationB' THEN RETURN; END_IF;
    IF "FRK_PersistImages".D013.Ordinal <> 1 THEN RETURN; END_IF;
    IF "FRK_PersistImages".D013.Payload.Info.Used THEN
        "FRK_SetRuntime".Work[2].Payload := "FRK_PersistImages".D013.Payload;
        IF NOT "FRK_SetShape"(RootIndex := 2, RootIdentity := 'StationB') THEN RETURN; END_IF;
    END_IF;
    "FRK_SetStore".Sets[2, 1] := "FRK_PersistImages".D013.Payload;
    "FRK_SetStore".SchemaVersion := 1;
    #FRK_DocApply_D013 := TRUE;
END_FUNCTION
FUNCTION "FRK_DocCapture_D014" : Bool
{ S7_Optimized_Access := 'TRUE' }
VERSION : 0.1
VAR_IN_OUT
    Length : DInt;
END_VAR
VAR_TEMP
    Index : Int;
    Stored : Int;
    Position : DInt;
    NativeResult : Int;
    Ok : Bool;
END_VAR
BEGIN
    #FRK_DocCapture_D014 := FALSE;
    "FRK_PersistImages".D014.SchemaVersion := 1; "FRK_PersistImages".D014.Scope := 'StationB';
    "FRK_PersistImages".D014.Ordinal := 2;
    "FRK_PersistImages".D014.Payload := "FRK_SetStore".Sets[2, 2];
    FOR #Index := 0 TO 9359 DO "FRK_PersistBuffers".D014Data[#Index] := BYTE#0; END_FOR;
    #Position := 24;
    #NativeResult := Serialize(SRC_VARIABLE := "FRK_PersistImages".D014, DEST_ARRAY => "FRK_PersistBuffers".D014Data, POS := #Position);
    IF #NativeResult <> 0 OR #Position < 24 OR #Position > 9360 THEN RETURN; END_IF;
    #Length := #Position - 24;
    #FRK_DocCapture_D014 := TRUE;
END_FUNCTION
FUNCTION "FRK_DocApply_D014" : Bool
{ S7_Optimized_Access := 'TRUE' }
VERSION : 0.1
VAR_TEMP
    Index : Int;
    Stored : Int;
    Position : DInt;
    NativeResult : Int;
    Ok : Bool;
END_VAR
BEGIN
    #FRK_DocApply_D014 := FALSE;
    #Position := 24;
    #NativeResult := Deserialize(SRC_ARRAY := "FRK_PersistBuffers".D014Data, DEST_VARIABLE => "FRK_PersistImages".D014, POS := #Position);
    IF #NativeResult <> 0 OR #Position <> 24 + UDINT_TO_DINT("FRK_PersistConsumers".Rows[14].Result.Length) THEN RETURN; END_IF;
    IF "FRK_PersistImages".D014.SchemaVersion <> 1 OR "FRK_PersistImages".D014.Scope <> 'StationB' THEN RETURN; END_IF;
    IF "FRK_PersistImages".D014.Ordinal <> 2 THEN RETURN; END_IF;
    IF "FRK_PersistImages".D014.Payload.Info.Used THEN
        "FRK_SetRuntime".Work[2].Payload := "FRK_PersistImages".D014.Payload;
        IF NOT "FRK_SetShape"(RootIndex := 2, RootIdentity := 'StationB') THEN RETURN; END_IF;
    END_IF;
    "FRK_SetStore".Sets[2, 2] := "FRK_PersistImages".D014.Payload;
    "FRK_SetStore".SchemaVersion := 1;
    #FRK_DocApply_D014 := TRUE;
END_FUNCTION
FUNCTION "FRK_DocCapture_D015" : Bool
{ S7_Optimized_Access := 'TRUE' }
VERSION : 0.1
VAR_IN_OUT
    Length : DInt;
END_VAR
VAR_TEMP
    Index : Int;
    Stored : Int;
    Position : DInt;
    NativeResult : Int;
    Ok : Bool;
END_VAR
BEGIN
    #FRK_DocCapture_D015 := FALSE;
    "FRK_PersistImages".D015.SchemaVersion := 1; "FRK_PersistImages".D015.Scope := 'StationB';
    "FRK_PersistImages".D015.Ordinal := 3;
    "FRK_PersistImages".D015.Payload := "FRK_SetStore".Sets[2, 3];
    FOR #Index := 0 TO 9359 DO "FRK_PersistBuffers".D015Data[#Index] := BYTE#0; END_FOR;
    #Position := 24;
    #NativeResult := Serialize(SRC_VARIABLE := "FRK_PersistImages".D015, DEST_ARRAY => "FRK_PersistBuffers".D015Data, POS := #Position);
    IF #NativeResult <> 0 OR #Position < 24 OR #Position > 9360 THEN RETURN; END_IF;
    #Length := #Position - 24;
    #FRK_DocCapture_D015 := TRUE;
END_FUNCTION
FUNCTION "FRK_DocApply_D015" : Bool
{ S7_Optimized_Access := 'TRUE' }
VERSION : 0.1
VAR_TEMP
    Index : Int;
    Stored : Int;
    Position : DInt;
    NativeResult : Int;
    Ok : Bool;
END_VAR
BEGIN
    #FRK_DocApply_D015 := FALSE;
    #Position := 24;
    #NativeResult := Deserialize(SRC_ARRAY := "FRK_PersistBuffers".D015Data, DEST_VARIABLE => "FRK_PersistImages".D015, POS := #Position);
    IF #NativeResult <> 0 OR #Position <> 24 + UDINT_TO_DINT("FRK_PersistConsumers".Rows[15].Result.Length) THEN RETURN; END_IF;
    IF "FRK_PersistImages".D015.SchemaVersion <> 1 OR "FRK_PersistImages".D015.Scope <> 'StationB' THEN RETURN; END_IF;
    IF "FRK_PersistImages".D015.Ordinal <> 3 THEN RETURN; END_IF;
    IF "FRK_PersistImages".D015.Payload.Info.Used THEN
        "FRK_SetRuntime".Work[2].Payload := "FRK_PersistImages".D015.Payload;
        IF NOT "FRK_SetShape"(RootIndex := 2, RootIdentity := 'StationB') THEN RETURN; END_IF;
    END_IF;
    "FRK_SetStore".Sets[2, 3] := "FRK_PersistImages".D015.Payload;
    "FRK_SetStore".SchemaVersion := 1;
    #FRK_DocApply_D015 := TRUE;
END_FUNCTION
FUNCTION "FRK_DocCapture_D016" : Bool
{ S7_Optimized_Access := 'TRUE' }
VERSION : 0.1
VAR_IN_OUT
    Length : DInt;
END_VAR
VAR_TEMP
    Index : Int;
    Stored : Int;
    Position : DInt;
    NativeResult : Int;
    Ok : Bool;
END_VAR
BEGIN
    #FRK_DocCapture_D016 := FALSE;
    "FRK_PersistImages".D016.SchemaVersion := 1; "FRK_PersistImages".D016.Scope := 'StationB';
    "FRK_PersistImages".D016.Ordinal := 4;
    "FRK_PersistImages".D016.Payload := "FRK_SetStore".Sets[2, 4];
    FOR #Index := 0 TO 9359 DO "FRK_PersistBuffers".D016Data[#Index] := BYTE#0; END_FOR;
    #Position := 24;
    #NativeResult := Serialize(SRC_VARIABLE := "FRK_PersistImages".D016, DEST_ARRAY => "FRK_PersistBuffers".D016Data, POS := #Position);
    IF #NativeResult <> 0 OR #Position < 24 OR #Position > 9360 THEN RETURN; END_IF;
    #Length := #Position - 24;
    #FRK_DocCapture_D016 := TRUE;
END_FUNCTION
FUNCTION "FRK_DocApply_D016" : Bool
{ S7_Optimized_Access := 'TRUE' }
VERSION : 0.1
VAR_TEMP
    Index : Int;
    Stored : Int;
    Position : DInt;
    NativeResult : Int;
    Ok : Bool;
END_VAR
BEGIN
    #FRK_DocApply_D016 := FALSE;
    #Position := 24;
    #NativeResult := Deserialize(SRC_ARRAY := "FRK_PersistBuffers".D016Data, DEST_VARIABLE => "FRK_PersistImages".D016, POS := #Position);
    IF #NativeResult <> 0 OR #Position <> 24 + UDINT_TO_DINT("FRK_PersistConsumers".Rows[16].Result.Length) THEN RETURN; END_IF;
    IF "FRK_PersistImages".D016.SchemaVersion <> 1 OR "FRK_PersistImages".D016.Scope <> 'StationB' THEN RETURN; END_IF;
    IF "FRK_PersistImages".D016.Ordinal <> 4 THEN RETURN; END_IF;
    IF "FRK_PersistImages".D016.Payload.Info.Used THEN
        "FRK_SetRuntime".Work[2].Payload := "FRK_PersistImages".D016.Payload;
        IF NOT "FRK_SetShape"(RootIndex := 2, RootIdentity := 'StationB') THEN RETURN; END_IF;
    END_IF;
    "FRK_SetStore".Sets[2, 4] := "FRK_PersistImages".D016.Payload;
    "FRK_SetStore".SchemaVersion := 1;
    #FRK_DocApply_D016 := TRUE;
END_FUNCTION
FUNCTION "FRK_DocCapture_D017" : Bool
{ S7_Optimized_Access := 'TRUE' }
VERSION : 0.1
VAR_IN_OUT
    Length : DInt;
END_VAR
VAR_TEMP
    Index : Int;
    Stored : Int;
    Position : DInt;
    NativeResult : Int;
    Ok : Bool;
END_VAR
BEGIN
    #FRK_DocCapture_D017 := FALSE;
    "FRK_PersistImages".D017.SchemaVersion := 1; "FRK_PersistImages".D017.Scope := 'users';
    IF NOT "FRK_AccessStorage".UsersReady THEN RETURN; END_IF;
    "FRK_PersistImages".D017.Generation := "FRK_LocalUsers".Generation;
    "FRK_PersistImages".D017.Count := "FRK_LocalUsers".Count;
    "FRK_PersistImages".D017.Rows := "FRK_LocalUsers".Rows;
    "FRK_PersistImages".D017.Checksum := "FRK_LocalUsers".Checksum;
    FOR #Index := 0 TO 8727 DO "FRK_PersistBuffers".D017Data[#Index] := BYTE#0; END_FOR;
    #Position := 24;
    #NativeResult := Serialize(SRC_VARIABLE := "FRK_PersistImages".D017, DEST_ARRAY => "FRK_PersistBuffers".D017Data, POS := #Position);
    IF #NativeResult <> 0 OR #Position < 24 OR #Position > 8728 THEN RETURN; END_IF;
    #Length := #Position - 24;
    #FRK_DocCapture_D017 := TRUE;
END_FUNCTION
FUNCTION "FRK_DocApply_D017" : Bool
{ S7_Optimized_Access := 'TRUE' }
VERSION : 0.1
VAR_TEMP
    Index : Int;
    Stored : Int;
    Position : DInt;
    NativeResult : Int;
    Ok : Bool;
END_VAR
BEGIN
    #FRK_DocApply_D017 := FALSE;
    #Position := 24;
    #NativeResult := Deserialize(SRC_ARRAY := "FRK_PersistBuffers".D017Data, DEST_VARIABLE => "FRK_PersistImages".D017, POS := #Position);
    IF #NativeResult <> 0 OR #Position <> 24 + UDINT_TO_DINT("FRK_PersistConsumers".Rows[17].Result.Length) THEN RETURN; END_IF;
    IF "FRK_PersistImages".D017.SchemaVersion <> 1 OR "FRK_PersistImages".D017.Scope <> 'users' THEN RETURN; END_IF;
    IF "FRK_PersistImages".D017.Generation = 0 OR NOT "FRK_AccessUsersShapeData"(Count := "FRK_PersistImages".D017.Count, Rows := "FRK_PersistImages".D017.Rows) THEN RETURN; END_IF;
    IF "FRK_PersistImages".D017.Checksum <> "FRK_AccessUsersCrcData"(SchemaVersion := "FRK_PersistImages".D017.SchemaVersion, Generation := "FRK_PersistImages".D017.Generation, Count := "FRK_PersistImages".D017.Count, Rows := "FRK_PersistImages".D017.Rows) THEN RETURN; END_IF;
    "FRK_LocalUsers".Generation := "FRK_PersistImages".D017.Generation;
    "FRK_LocalUsers".Count := "FRK_PersistImages".D017.Count;
    "FRK_LocalUsers".Rows := "FRK_PersistImages".D017.Rows;
    "FRK_LocalUsers".Checksum := "FRK_PersistImages".D017.Checksum;
    "FRK_LocalUsers".SchemaVersion := 1; "FRK_AccessStorage".UsersCommissioned := TRUE;
    #FRK_DocApply_D017 := TRUE;
END_FUNCTION
FUNCTION "FRK_DocReject" : Void
{ S7_Optimized_Access := 'TRUE' }
VERSION : 0.1
VAR_INPUT
    Slot : Int;
END_VAR
VAR_TEMP
    Stored : Int;
END_VAR
BEGIN
    CASE #Slot OF
        1:
            #Stored := "FRK_ConfigFind"(Scope := 'StationA', Key := 'siteLabel', ModelCode := '');
            IF #Stored > 0 THEN "FRK_ConfigStore".Rows[#Stored].Used := FALSE; END_IF;
            #Stored := "FRK_ConfigFind"(Scope := 'StationA', Key := 'long.kkkkkkkkkkkkkkkkkkkkkkkkkkkkkkkkkkkkkkkkkkkkkkkkkkkkkkkkkkkkkkkkkkkkkkkkkkkkkkkkkkkkkkkkkkkkkkkkkkkkkkkkkkkkkkkkkkkkkkkkkkkkkkkkkkkkkkk', ModelCode := '');
            IF #Stored > 0 THEN "FRK_ConfigStore".Rows[#Stored].Used := FALSE; END_IF;
            #Stored := "FRK_ConfigFind"(Scope := 'StationA', Key := 'enabled', ModelCode := '');
            IF #Stored > 0 THEN "FRK_ConfigStore".Rows[#Stored].Used := FALSE; END_IF;
            #Stored := "FRK_ConfigFind"(Scope := 'StationA.Satellite', Key := 'siteLabel', ModelCode := '');
            IF #Stored > 0 THEN "FRK_ConfigStore".Rows[#Stored].Used := FALSE; END_IF;
            #Stored := "FRK_ConfigFind"(Scope := 'StationA.Satellite', Key := 'long.kkkkkkkkkkkkkkkkkkkkkkkkkkkkkkkkkkkkkkkkkkkkkkkkkkkkkkkkkkkkkkkkkkkkkkkkkkkkkkkkkkkkkkkkkkkkkkkkkkkkkkkkkkkkkkkkkkkkkkkkkkkkkkkkkkkkkkk', ModelCode := '');
            IF #Stored > 0 THEN "FRK_ConfigStore".Rows[#Stored].Used := FALSE; END_IF;
            #Stored := "FRK_ConfigFind"(Scope := 'StationA.Satellite', Key := 'enabled', ModelCode := '');
            IF #Stored > 0 THEN "FRK_ConfigStore".Rows[#Stored].Used := FALSE; END_IF;
            #Stored := "FRK_ConfigFind"(Scope := 'StationA.Satellite.Inner', Key := 'siteLabel', ModelCode := '');
            IF #Stored > 0 THEN "FRK_ConfigStore".Rows[#Stored].Used := FALSE; END_IF;
            #Stored := "FRK_ConfigFind"(Scope := 'StationA.Satellite.Inner', Key := 'long.kkkkkkkkkkkkkkkkkkkkkkkkkkkkkkkkkkkkkkkkkkkkkkkkkkkkkkkkkkkkkkkkkkkkkkkkkkkkkkkkkkkkkkkkkkkkkkkkkkkkkkkkkkkkkkkkkkkkkkkkkkkkkkkkkkkkkkk', ModelCode := '');
            IF #Stored > 0 THEN "FRK_ConfigStore".Rows[#Stored].Used := FALSE; END_IF;
            #Stored := "FRK_ConfigFind"(Scope := 'StationA.Satellite.Inner', Key := 'enabled', ModelCode := '');
            IF #Stored > 0 THEN "FRK_ConfigStore".Rows[#Stored].Used := FALSE; END_IF;
            "FRK_ConfigLoss"(RootIndex := 1, Scope := 'StationA');
        2:
            #Stored := "FRK_ConfigFind"(Scope := 'StationA', Key := 'timeout', ModelCode := 'MODEL_A');
            IF #Stored > 0 THEN "FRK_ConfigStore".Rows[#Stored].Used := FALSE; END_IF;
            #Stored := "FRK_ConfigFind"(Scope := 'StationA', Key := 'preset', ModelCode := 'MODEL_A');
            IF #Stored > 0 THEN "FRK_ConfigStore".Rows[#Stored].Used := FALSE; END_IF;
            #Stored := "FRK_ConfigFind"(Scope := 'StationA.Cell', Key := 'timeout', ModelCode := 'MODEL_A');
            IF #Stored > 0 THEN "FRK_ConfigStore".Rows[#Stored].Used := FALSE; END_IF;
            #Stored := "FRK_ConfigFind"(Scope := 'StationA.Cell', Key := 'preset', ModelCode := 'MODEL_A');
            IF #Stored > 0 THEN "FRK_ConfigStore".Rows[#Stored].Used := FALSE; END_IF;
            #Stored := "FRK_ConfigFind"(Scope := 'StationA.Cell.Clamp', Key := 'timeout', ModelCode := 'MODEL_A');
            IF #Stored > 0 THEN "FRK_ConfigStore".Rows[#Stored].Used := FALSE; END_IF;
            #Stored := "FRK_ConfigFind"(Scope := 'StationA.Cell.Clamp', Key := 'preset', ModelCode := 'MODEL_A');
            IF #Stored > 0 THEN "FRK_ConfigStore".Rows[#Stored].Used := FALSE; END_IF;
            #Stored := "FRK_ConfigFind"(Scope := 'StationA.Cell.Gate', Key := 'timeout', ModelCode := 'MODEL_A');
            IF #Stored > 0 THEN "FRK_ConfigStore".Rows[#Stored].Used := FALSE; END_IF;
            #Stored := "FRK_ConfigFind"(Scope := 'StationA.Cell.Gate', Key := 'preset', ModelCode := 'MODEL_A');
            IF #Stored > 0 THEN "FRK_ConfigStore".Rows[#Stored].Used := FALSE; END_IF;
            #Stored := "FRK_ConfigFind"(Scope := 'StationA.Satellite', Key := 'timeout', ModelCode := 'MODEL_A');
            IF #Stored > 0 THEN "FRK_ConfigStore".Rows[#Stored].Used := FALSE; END_IF;
            #Stored := "FRK_ConfigFind"(Scope := 'StationA.Satellite', Key := 'preset', ModelCode := 'MODEL_A');
            IF #Stored > 0 THEN "FRK_ConfigStore".Rows[#Stored].Used := FALSE; END_IF;
            #Stored := "FRK_ConfigFind"(Scope := 'StationA.Satellite.Cell', Key := 'timeout', ModelCode := 'MODEL_A');
            IF #Stored > 0 THEN "FRK_ConfigStore".Rows[#Stored].Used := FALSE; END_IF;
            #Stored := "FRK_ConfigFind"(Scope := 'StationA.Satellite.Cell', Key := 'preset', ModelCode := 'MODEL_A');
            IF #Stored > 0 THEN "FRK_ConfigStore".Rows[#Stored].Used := FALSE; END_IF;
            #Stored := "FRK_ConfigFind"(Scope := 'StationA.Satellite.Cell.Clamp', Key := 'timeout', ModelCode := 'MODEL_A');
            IF #Stored > 0 THEN "FRK_ConfigStore".Rows[#Stored].Used := FALSE; END_IF;
            #Stored := "FRK_ConfigFind"(Scope := 'StationA.Satellite.Cell.Clamp', Key := 'preset', ModelCode := 'MODEL_A');
            IF #Stored > 0 THEN "FRK_ConfigStore".Rows[#Stored].Used := FALSE; END_IF;
            #Stored := "FRK_ConfigFind"(Scope := 'StationA.Satellite.Cell.Gate', Key := 'timeout', ModelCode := 'MODEL_A');
            IF #Stored > 0 THEN "FRK_ConfigStore".Rows[#Stored].Used := FALSE; END_IF;
            #Stored := "FRK_ConfigFind"(Scope := 'StationA.Satellite.Cell.Gate', Key := 'preset', ModelCode := 'MODEL_A');
            IF #Stored > 0 THEN "FRK_ConfigStore".Rows[#Stored].Used := FALSE; END_IF;
            #Stored := "FRK_ConfigFind"(Scope := 'StationA.Satellite.Inner', Key := 'timeout', ModelCode := 'MODEL_A');
            IF #Stored > 0 THEN "FRK_ConfigStore".Rows[#Stored].Used := FALSE; END_IF;
            #Stored := "FRK_ConfigFind"(Scope := 'StationA.Satellite.Inner', Key := 'preset', ModelCode := 'MODEL_A');
            IF #Stored > 0 THEN "FRK_ConfigStore".Rows[#Stored].Used := FALSE; END_IF;
            #Stored := "FRK_ConfigFind"(Scope := 'StationA.Satellite.Inner.Cell', Key := 'timeout', ModelCode := 'MODEL_A');
            IF #Stored > 0 THEN "FRK_ConfigStore".Rows[#Stored].Used := FALSE; END_IF;
            #Stored := "FRK_ConfigFind"(Scope := 'StationA.Satellite.Inner.Cell', Key := 'preset', ModelCode := 'MODEL_A');
            IF #Stored > 0 THEN "FRK_ConfigStore".Rows[#Stored].Used := FALSE; END_IF;
            #Stored := "FRK_ConfigFind"(Scope := 'StationA.Satellite.Inner.Cell.Clamp', Key := 'timeout', ModelCode := 'MODEL_A');
            IF #Stored > 0 THEN "FRK_ConfigStore".Rows[#Stored].Used := FALSE; END_IF;
            #Stored := "FRK_ConfigFind"(Scope := 'StationA.Satellite.Inner.Cell.Clamp', Key := 'preset', ModelCode := 'MODEL_A');
            IF #Stored > 0 THEN "FRK_ConfigStore".Rows[#Stored].Used := FALSE; END_IF;
            #Stored := "FRK_ConfigFind"(Scope := 'StationA.Satellite.Inner.Cell.Gate', Key := 'timeout', ModelCode := 'MODEL_A');
            IF #Stored > 0 THEN "FRK_ConfigStore".Rows[#Stored].Used := FALSE; END_IF;
            #Stored := "FRK_ConfigFind"(Scope := 'StationA.Satellite.Inner.Cell.Gate', Key := 'preset', ModelCode := 'MODEL_A');
            IF #Stored > 0 THEN "FRK_ConfigStore".Rows[#Stored].Used := FALSE; END_IF;
            "FRK_ConfigLoss"(RootIndex := 1, Scope := 'StationA');
        3:
            #Stored := "FRK_ConfigFind"(Scope := 'StationA', Key := 'timeout', ModelCode := 'MODEL_B');
            IF #Stored > 0 THEN "FRK_ConfigStore".Rows[#Stored].Used := FALSE; END_IF;
            #Stored := "FRK_ConfigFind"(Scope := 'StationA', Key := 'preset', ModelCode := 'MODEL_B');
            IF #Stored > 0 THEN "FRK_ConfigStore".Rows[#Stored].Used := FALSE; END_IF;
            #Stored := "FRK_ConfigFind"(Scope := 'StationA.Cell', Key := 'timeout', ModelCode := 'MODEL_B');
            IF #Stored > 0 THEN "FRK_ConfigStore".Rows[#Stored].Used := FALSE; END_IF;
            #Stored := "FRK_ConfigFind"(Scope := 'StationA.Cell', Key := 'preset', ModelCode := 'MODEL_B');
            IF #Stored > 0 THEN "FRK_ConfigStore".Rows[#Stored].Used := FALSE; END_IF;
            #Stored := "FRK_ConfigFind"(Scope := 'StationA.Cell.Clamp', Key := 'timeout', ModelCode := 'MODEL_B');
            IF #Stored > 0 THEN "FRK_ConfigStore".Rows[#Stored].Used := FALSE; END_IF;
            #Stored := "FRK_ConfigFind"(Scope := 'StationA.Cell.Clamp', Key := 'preset', ModelCode := 'MODEL_B');
            IF #Stored > 0 THEN "FRK_ConfigStore".Rows[#Stored].Used := FALSE; END_IF;
            #Stored := "FRK_ConfigFind"(Scope := 'StationA.Cell.Gate', Key := 'timeout', ModelCode := 'MODEL_B');
            IF #Stored > 0 THEN "FRK_ConfigStore".Rows[#Stored].Used := FALSE; END_IF;
            #Stored := "FRK_ConfigFind"(Scope := 'StationA.Cell.Gate', Key := 'preset', ModelCode := 'MODEL_B');
            IF #Stored > 0 THEN "FRK_ConfigStore".Rows[#Stored].Used := FALSE; END_IF;
            #Stored := "FRK_ConfigFind"(Scope := 'StationA.Satellite', Key := 'timeout', ModelCode := 'MODEL_B');
            IF #Stored > 0 THEN "FRK_ConfigStore".Rows[#Stored].Used := FALSE; END_IF;
            #Stored := "FRK_ConfigFind"(Scope := 'StationA.Satellite', Key := 'preset', ModelCode := 'MODEL_B');
            IF #Stored > 0 THEN "FRK_ConfigStore".Rows[#Stored].Used := FALSE; END_IF;
            #Stored := "FRK_ConfigFind"(Scope := 'StationA.Satellite.Cell', Key := 'timeout', ModelCode := 'MODEL_B');
            IF #Stored > 0 THEN "FRK_ConfigStore".Rows[#Stored].Used := FALSE; END_IF;
            #Stored := "FRK_ConfigFind"(Scope := 'StationA.Satellite.Cell', Key := 'preset', ModelCode := 'MODEL_B');
            IF #Stored > 0 THEN "FRK_ConfigStore".Rows[#Stored].Used := FALSE; END_IF;
            #Stored := "FRK_ConfigFind"(Scope := 'StationA.Satellite.Cell.Clamp', Key := 'timeout', ModelCode := 'MODEL_B');
            IF #Stored > 0 THEN "FRK_ConfigStore".Rows[#Stored].Used := FALSE; END_IF;
            #Stored := "FRK_ConfigFind"(Scope := 'StationA.Satellite.Cell.Clamp', Key := 'preset', ModelCode := 'MODEL_B');
            IF #Stored > 0 THEN "FRK_ConfigStore".Rows[#Stored].Used := FALSE; END_IF;
            #Stored := "FRK_ConfigFind"(Scope := 'StationA.Satellite.Cell.Gate', Key := 'timeout', ModelCode := 'MODEL_B');
            IF #Stored > 0 THEN "FRK_ConfigStore".Rows[#Stored].Used := FALSE; END_IF;
            #Stored := "FRK_ConfigFind"(Scope := 'StationA.Satellite.Cell.Gate', Key := 'preset', ModelCode := 'MODEL_B');
            IF #Stored > 0 THEN "FRK_ConfigStore".Rows[#Stored].Used := FALSE; END_IF;
            #Stored := "FRK_ConfigFind"(Scope := 'StationA.Satellite.Inner', Key := 'timeout', ModelCode := 'MODEL_B');
            IF #Stored > 0 THEN "FRK_ConfigStore".Rows[#Stored].Used := FALSE; END_IF;
            #Stored := "FRK_ConfigFind"(Scope := 'StationA.Satellite.Inner', Key := 'preset', ModelCode := 'MODEL_B');
            IF #Stored > 0 THEN "FRK_ConfigStore".Rows[#Stored].Used := FALSE; END_IF;
            #Stored := "FRK_ConfigFind"(Scope := 'StationA.Satellite.Inner.Cell', Key := 'timeout', ModelCode := 'MODEL_B');
            IF #Stored > 0 THEN "FRK_ConfigStore".Rows[#Stored].Used := FALSE; END_IF;
            #Stored := "FRK_ConfigFind"(Scope := 'StationA.Satellite.Inner.Cell', Key := 'preset', ModelCode := 'MODEL_B');
            IF #Stored > 0 THEN "FRK_ConfigStore".Rows[#Stored].Used := FALSE; END_IF;
            #Stored := "FRK_ConfigFind"(Scope := 'StationA.Satellite.Inner.Cell.Clamp', Key := 'timeout', ModelCode := 'MODEL_B');
            IF #Stored > 0 THEN "FRK_ConfigStore".Rows[#Stored].Used := FALSE; END_IF;
            #Stored := "FRK_ConfigFind"(Scope := 'StationA.Satellite.Inner.Cell.Clamp', Key := 'preset', ModelCode := 'MODEL_B');
            IF #Stored > 0 THEN "FRK_ConfigStore".Rows[#Stored].Used := FALSE; END_IF;
            #Stored := "FRK_ConfigFind"(Scope := 'StationA.Satellite.Inner.Cell.Gate', Key := 'timeout', ModelCode := 'MODEL_B');
            IF #Stored > 0 THEN "FRK_ConfigStore".Rows[#Stored].Used := FALSE; END_IF;
            #Stored := "FRK_ConfigFind"(Scope := 'StationA.Satellite.Inner.Cell.Gate', Key := 'preset', ModelCode := 'MODEL_B');
            IF #Stored > 0 THEN "FRK_ConfigStore".Rows[#Stored].Used := FALSE; END_IF;
            "FRK_ConfigLoss"(RootIndex := 1, Scope := 'StationA');
        4:
            "FRK_AccessPolicies".Rows[1].Scope := 'StationA';
            "FRK_AccessPolicies".Rows[1].SchemaVersion := 0;
            "FRK_AccessPolicies".Rows[1].Initialized := TRUE;
        5:
            "FRK_SetStore".Sets[1, 1].Info.Used := FALSE;
            "FRK_ConfigLoss"(RootIndex := 1, Scope := 'StationA');
        6:
            "FRK_SetStore".Sets[1, 2].Info.Used := FALSE;
            "FRK_ConfigLoss"(RootIndex := 1, Scope := 'StationA');
        7:
            "FRK_SetStore".Sets[1, 3].Info.Used := FALSE;
            "FRK_ConfigLoss"(RootIndex := 1, Scope := 'StationA');
        8:
            "FRK_SetStore".Sets[1, 4].Info.Used := FALSE;
            "FRK_ConfigLoss"(RootIndex := 1, Scope := 'StationA');
        9:
            #Stored := "FRK_ConfigFind"(Scope := 'StationB', Key := 'siteLabel', ModelCode := '');
            IF #Stored > 0 THEN "FRK_ConfigStore".Rows[#Stored].Used := FALSE; END_IF;
            #Stored := "FRK_ConfigFind"(Scope := 'StationB', Key := 'long.kkkkkkkkkkkkkkkkkkkkkkkkkkkkkkkkkkkkkkkkkkkkkkkkkkkkkkkkkkkkkkkkkkkkkkkkkkkkkkkkkkkkkkkkkkkkkkkkkkkkkkkkkkkkkkkkkkkkkkkkkkkkkkkkkkkkkkk', ModelCode := '');
            IF #Stored > 0 THEN "FRK_ConfigStore".Rows[#Stored].Used := FALSE; END_IF;
            #Stored := "FRK_ConfigFind"(Scope := 'StationB', Key := 'enabled', ModelCode := '');
            IF #Stored > 0 THEN "FRK_ConfigStore".Rows[#Stored].Used := FALSE; END_IF;
            #Stored := "FRK_ConfigFind"(Scope := 'StationB.Satellite', Key := 'siteLabel', ModelCode := '');
            IF #Stored > 0 THEN "FRK_ConfigStore".Rows[#Stored].Used := FALSE; END_IF;
            #Stored := "FRK_ConfigFind"(Scope := 'StationB.Satellite', Key := 'long.kkkkkkkkkkkkkkkkkkkkkkkkkkkkkkkkkkkkkkkkkkkkkkkkkkkkkkkkkkkkkkkkkkkkkkkkkkkkkkkkkkkkkkkkkkkkkkkkkkkkkkkkkkkkkkkkkkkkkkkkkkkkkkkkkkkkkkk', ModelCode := '');
            IF #Stored > 0 THEN "FRK_ConfigStore".Rows[#Stored].Used := FALSE; END_IF;
            #Stored := "FRK_ConfigFind"(Scope := 'StationB.Satellite', Key := 'enabled', ModelCode := '');
            IF #Stored > 0 THEN "FRK_ConfigStore".Rows[#Stored].Used := FALSE; END_IF;
            #Stored := "FRK_ConfigFind"(Scope := 'StationB.Satellite.Inner', Key := 'siteLabel', ModelCode := '');
            IF #Stored > 0 THEN "FRK_ConfigStore".Rows[#Stored].Used := FALSE; END_IF;
            #Stored := "FRK_ConfigFind"(Scope := 'StationB.Satellite.Inner', Key := 'long.kkkkkkkkkkkkkkkkkkkkkkkkkkkkkkkkkkkkkkkkkkkkkkkkkkkkkkkkkkkkkkkkkkkkkkkkkkkkkkkkkkkkkkkkkkkkkkkkkkkkkkkkkkkkkkkkkkkkkkkkkkkkkkkkkkkkkkk', ModelCode := '');
            IF #Stored > 0 THEN "FRK_ConfigStore".Rows[#Stored].Used := FALSE; END_IF;
            #Stored := "FRK_ConfigFind"(Scope := 'StationB.Satellite.Inner', Key := 'enabled', ModelCode := '');
            IF #Stored > 0 THEN "FRK_ConfigStore".Rows[#Stored].Used := FALSE; END_IF;
            "FRK_ConfigLoss"(RootIndex := 2, Scope := 'StationB');
        10:
            #Stored := "FRK_ConfigFind"(Scope := 'StationB', Key := 'timeout', ModelCode := 'MODEL_A');
            IF #Stored > 0 THEN "FRK_ConfigStore".Rows[#Stored].Used := FALSE; END_IF;
            #Stored := "FRK_ConfigFind"(Scope := 'StationB', Key := 'preset', ModelCode := 'MODEL_A');
            IF #Stored > 0 THEN "FRK_ConfigStore".Rows[#Stored].Used := FALSE; END_IF;
            #Stored := "FRK_ConfigFind"(Scope := 'StationB.Cell', Key := 'timeout', ModelCode := 'MODEL_A');
            IF #Stored > 0 THEN "FRK_ConfigStore".Rows[#Stored].Used := FALSE; END_IF;
            #Stored := "FRK_ConfigFind"(Scope := 'StationB.Cell', Key := 'preset', ModelCode := 'MODEL_A');
            IF #Stored > 0 THEN "FRK_ConfigStore".Rows[#Stored].Used := FALSE; END_IF;
            #Stored := "FRK_ConfigFind"(Scope := 'StationB.Cell.Clamp', Key := 'timeout', ModelCode := 'MODEL_A');
            IF #Stored > 0 THEN "FRK_ConfigStore".Rows[#Stored].Used := FALSE; END_IF;
            #Stored := "FRK_ConfigFind"(Scope := 'StationB.Cell.Clamp', Key := 'preset', ModelCode := 'MODEL_A');
            IF #Stored > 0 THEN "FRK_ConfigStore".Rows[#Stored].Used := FALSE; END_IF;
            #Stored := "FRK_ConfigFind"(Scope := 'StationB.Cell.Gate', Key := 'timeout', ModelCode := 'MODEL_A');
            IF #Stored > 0 THEN "FRK_ConfigStore".Rows[#Stored].Used := FALSE; END_IF;
            #Stored := "FRK_ConfigFind"(Scope := 'StationB.Cell.Gate', Key := 'preset', ModelCode := 'MODEL_A');
            IF #Stored > 0 THEN "FRK_ConfigStore".Rows[#Stored].Used := FALSE; END_IF;
            #Stored := "FRK_ConfigFind"(Scope := 'StationB.Satellite', Key := 'timeout', ModelCode := 'MODEL_A');
            IF #Stored > 0 THEN "FRK_ConfigStore".Rows[#Stored].Used := FALSE; END_IF;
            #Stored := "FRK_ConfigFind"(Scope := 'StationB.Satellite', Key := 'preset', ModelCode := 'MODEL_A');
            IF #Stored > 0 THEN "FRK_ConfigStore".Rows[#Stored].Used := FALSE; END_IF;
            #Stored := "FRK_ConfigFind"(Scope := 'StationB.Satellite.Cell', Key := 'timeout', ModelCode := 'MODEL_A');
            IF #Stored > 0 THEN "FRK_ConfigStore".Rows[#Stored].Used := FALSE; END_IF;
            #Stored := "FRK_ConfigFind"(Scope := 'StationB.Satellite.Cell', Key := 'preset', ModelCode := 'MODEL_A');
            IF #Stored > 0 THEN "FRK_ConfigStore".Rows[#Stored].Used := FALSE; END_IF;
            #Stored := "FRK_ConfigFind"(Scope := 'StationB.Satellite.Cell.Clamp', Key := 'timeout', ModelCode := 'MODEL_A');
            IF #Stored > 0 THEN "FRK_ConfigStore".Rows[#Stored].Used := FALSE; END_IF;
            #Stored := "FRK_ConfigFind"(Scope := 'StationB.Satellite.Cell.Clamp', Key := 'preset', ModelCode := 'MODEL_A');
            IF #Stored > 0 THEN "FRK_ConfigStore".Rows[#Stored].Used := FALSE; END_IF;
            #Stored := "FRK_ConfigFind"(Scope := 'StationB.Satellite.Cell.Gate', Key := 'timeout', ModelCode := 'MODEL_A');
            IF #Stored > 0 THEN "FRK_ConfigStore".Rows[#Stored].Used := FALSE; END_IF;
            #Stored := "FRK_ConfigFind"(Scope := 'StationB.Satellite.Cell.Gate', Key := 'preset', ModelCode := 'MODEL_A');
            IF #Stored > 0 THEN "FRK_ConfigStore".Rows[#Stored].Used := FALSE; END_IF;
            #Stored := "FRK_ConfigFind"(Scope := 'StationB.Satellite.Inner', Key := 'timeout', ModelCode := 'MODEL_A');
            IF #Stored > 0 THEN "FRK_ConfigStore".Rows[#Stored].Used := FALSE; END_IF;
            #Stored := "FRK_ConfigFind"(Scope := 'StationB.Satellite.Inner', Key := 'preset', ModelCode := 'MODEL_A');
            IF #Stored > 0 THEN "FRK_ConfigStore".Rows[#Stored].Used := FALSE; END_IF;
            #Stored := "FRK_ConfigFind"(Scope := 'StationB.Satellite.Inner.Cell', Key := 'timeout', ModelCode := 'MODEL_A');
            IF #Stored > 0 THEN "FRK_ConfigStore".Rows[#Stored].Used := FALSE; END_IF;
